(* IEC 61131-3 sources: daoli-st-library/DL_Process (part 35) *)

(* ---- FB_DL_FormationWeekPlan.st ---- *)
(*
  ==================================================================
  组件名 Component  : FB_DL_FormationWeekPlan
  分类   Category   : DL_Process
  版本   Version    : 1.0.0
  功能   Purpose    : 周计划窗（周序号闸 + 月窗闸双闸）。把日历日换算成「月内周
                      序号（1..5）」与「周内日序号（1..7）」，两个闸同时成立才算
                      计划窗开启：一 月窗闸 = 当日落在组态的月内生产窗区间；
                      二 周序号闸 = 当日所在周序号落在允许的周区间。
                      同时给出周内与月内剩余天数，供上层排产节拍使用。
  溯源   Origin     : 周序号 / 月窗双闸为通用排产窗语义；本件为 clean-room 实现，
                      仅借鉴来源分类与参数域组织（来源标签 roadmap-p2-weekplan），
                      道莅原创设计，未复制任何闭源代码行。
  平台   Platform   : 纯 IEC 61131-3（INT 整除与 MOD，除子为常量，无私有库）
  作者   Author     : 道莅代码库 · PLC 编程专家（R55）
  ------------------------------------------------------------------
  边界 Boundary     :
                      一 本件只判双闸与剩余天数，不生成工单、不判产量；
                      二 周序号按「月内第几周」口径（1 日为第 1 周第 1 日），非 ISO 周；
                      三 整除与取模的除子均为常量 7，且除前已把日序回钳到 1..31；
                      四 双闸任一不成立即关窗，关窗原因由两个独立布尔出口区分（R190）；
                      五 无全局变量、无外部变量声明、无物理地址寻址。
  输出契约 Output contract:
                      bMonthGateOk / bWeekGateOk 为两条独立闸的实时值，
                      bWindowOpen 仅在两条闸同时成立时为真（挂状态量）；
                      nWeekIdx 域 1..5，nDayInWeek 域 1..7，两者恒由回钳后的日序派生；
                      eCause 故障级成因与 bError 配对（R45），信息级永不置 bError。
  修订记录 Revision  :
    2026-11-20  v1.0.0  R55 首版（批 2 · 序号 9）
  ==================================================================
*)

TYPE E_DL_FwpCause :
(
    eNone       := 0,   // 无成因 / no cause
    eCfgIllegal := 1,   // 组态非法：年月日、窗界或周区间越域（故障级，与 bError 配对）/ illegal config, calendar, window bounds or week band out of domain
    eMonthGate  := 2,   // 月窗闸不成立（信息级）/ the monthly window gate does not hold, informational
    eWeekGate   := 3    // 周序号闸不成立（信息级）/ the week index gate does not hold, informational
);
END_TYPE

FUNCTION_BLOCK FB_DL_FormationWeekPlan
VAR_INPUT
    bEnable      : BOOL := TRUE;             // 使能，失能时关窗 [-] / enable, the window closes when disabled
    bReset       : BOOL := FALSE;           // 复位上升沿清故障锁存 [-] / reset rising edge clears the fault latch
    nYear        : INT := 2026;              // 当前年份 [年]，域 2000..2100 / current year [year], domain 2000 to 2100
    nMonth       : INT := 1;                 // 当前月份 [月]，域 1..12 / current month [month], domain 1 to 12
    nDayOfMonth  : INT := 1;                 // 当月第几日 [日]，域 1..31 / day of month [day], domain 1 to 31
    nWinStartDay : INT := 1;                 // 月生产窗起始日 [日] / monthly production window start day [day]
    nWinEndDay   : INT := 28;                // 月生产窗结束日 [日]，须不早于起始日 / monthly window end day, not earlier than the start
    nWeekFrom    : INT := 1;                 // 允许的周序号下限（月内第几周）[周]，域 1..5 / allowed week index floor, domain 1 to 5
    nWeekTo      : INT := 5;                 // 允许的周序号上限（月内第几周）[周]，域 1..5 / allowed week index ceiling, domain 1 to 5
END_VAR
VAR_OUTPUT
    bWindowOpen  : BOOL := FALSE;            // 双闸同时成立（计划窗开启）[-] / both gates hold, the planning window is open
    bMonthGateOk : BOOL := FALSE;            // 月窗闸实时值 [-] / monthly window gate live value
    bWeekGateOk  : BOOL := FALSE;            // 周序号闸实时值 [-] / week index gate live value
    nWeekIdx     : INT := 1;                 // 月内周序号 [周]，域 1..5 / week index within the month, domain 1 to 5
    nDayInWeek   : INT := 1;                 // 周内日序号 [日]，域 1..7 / day index within the week, domain 1 to 7
    nRemainInWeek: INT := 0;                 // 本周剩余天数（不跨月）[日] / remaining days this week, not crossing the month
    nRemainInMonth : INT := 0;               // 本月剩余天数 [日] / remaining days this month
    nPlanDays    : INT := 0;                 // 本窗剩余可排产天数（双闸内计数）[日] / remaining plannable days inside the window
    eCause       : E_DL_FwpCause := E_DL_FwpCause.eNone; // 成因出口 [枚举] / cause outlet [enum]
    bError       : BOOL := FALSE;            // 故障锁存标志 [-] / fault latch flag
END_VAR
VAR
    rtReset      : R_TRIG;                   // 复位沿检测，段 0 无条件刷新 / reset edge detector, refreshed unconditionally in segment zero
    _eFaultCause : E_DL_FwpCause := E_DL_FwpCause.eNone;  // 故障级成因，锁存至复位沿 / fault cause, latched until the reset edge
    _bFault      : BOOL := FALSE;            // 故障锁存位 [-] / fault latch bit
    _bInit       : BOOL := FALSE;            // 首扫初始化完成标志（R310）/ first scan initialisation flag
    _bCfgBad     : BOOL := FALSE;            // 组态非法判定 [-] / illegal configuration verdict
    _bMonthGate  : BOOL := FALSE;            // 月窗闸工作值 [-] / monthly window gate working value
    _bWeekGate   : BOOL := FALSE;            // 周序号闸工作值 [-] / week index gate working value
    _nDaysInMonth: INT := 30;                // 当月日历天数 [日] / calendar days of the current month [day]
    _nDay        : INT := 1;                 // 回钳后的当日序号 [日] / clamped day index [day]
    _nStart      : INT := 1;                 // 回钳后的窗起始日 [日] / clamped window start day [day]
    _nEnd        : INT := 1;                 // 回钳后的窗结束日 [日] / clamped window end day [day]
    _nWeekFrom   : INT := 1;                 // 回钳后的周序号下限 [周] / clamped week index floor [week]
    _nWeekTo     : INT := 5;                 // 回钳后的周序号上限 [周] / clamped week index ceiling [week]
    _nWeekIdx    : INT := 1;                 // 周序号工作值 [周] / week index working value [week]
    _nDayInWeek  : INT := 1;                 // 周内日序号工作值 [日] / day in week working value [day]
    _nRemainWeek : INT := 0;                 // 本周剩余天数工作值 [日] / remaining week days working value [day]
    _nRemainMonth: INT := 0;                 // 本月剩余天数工作值 [日] / remaining month days working value [day]
    _nPlanDays   : INT := 0;                 // 窗内剩余可排产天数工作值 [日] / remaining plannable days working value [day]
    _nScanDay    : INT := 1;                 // 窗内扫描用日序（自当日到窗末）[日] / scanning day index from today to the window end [day]
END_VAR
VAR CONSTANT
    DL_FWP_DAY_MAX   : INT := 31;            // 月内最大天数 [日] / maximum days within a month [day]
    DL_FWP_WEEK_N    : INT := 7;             // 一周日数，整除去子（常量非零）[日] / days per week, the division divisor as a non-zero constant [day]
    DL_FWP_WEEK_MAX  : INT := 5;             // 月内最大周序号 [周] / maximum week index within a month [week]
    DL_FWP_YEAR_MIN  : INT := 2000;          // 年份下限 [年] / year floor [year]
    DL_FWP_YEAR_MAX  : INT := 2100;          // 年份上限 [年] / year ceiling [year]
END_VAR

// 段 0｜复位沿无条件周期刷新（禁入分支）/ segment 0, unconditional refresh of the reset edge, never inside a branch
rtReset(CLK := bReset); // 复位沿无条件刷新 / unconditional refresh of the reset edge

// 段 1｜首扫初始化（R310）/ segment 1, first scan initialisation
IF NOT _bInit THEN // 首扫一拍 / the very first scan
    _bInit := TRUE; // 置首扫完成标志 / raise the first scan flag
    _bFault := FALSE; // 故障锁存清零 / clear the fault latch
    _eFaultCause := E_DL_FwpCause.eNone; // 故障级成因清零 / clear the fault cause
    _nWeekIdx := 1; // 周序号从第一周起 / the week index starts at one
    _nDayInWeek := 1; // 周内日序号从第一日起 / the day in week starts at one
END_IF

// 段 2｜复位沿作用域：清故障锁存与故障级成因（不动日历派生量）/ segment 2, reset edge scope
IF rtReset.Q THEN // 复位沿 / reset edge
    _bFault := FALSE; // 作用域一：清故障锁存 / scope one, clear the fault latch
    _eFaultCause := E_DL_FwpCause.eNone; // 作用域一：清故障级成因 / scope one, clear the fault cause
END_IF

// 段 3｜日历天数：闰年二月二十九日 / segment 3, calendar days with a leap February
_nDaysInMonth := 31; // 默认三十一日 / default thirty one days
CASE nMonth OF
1, 3, 5, 7, 8, 10, 12: // 大月 / long months
    _nDaysInMonth := 31; // 三十一日 / thirty one days
2: // 二月 / february
    IF ((nYear MOD 4) = 0) AND (((nYear MOD 100) <> 0) OR ((nYear MOD 400) = 0)) THEN // 闰年判据 / leap year criterion
        _nDaysInMonth := 29; // 闰年二十九日 / twenty nine days in a leap year
    ELSE
        _nDaysInMonth := 28; // 平年二十八日 / twenty eight days in a common year
    END_IF
4, 6, 9, 11: // 小月 / short months
    _nDaysInMonth := 30; // 三十日 / thirty days
ELSE // 非法月份兜底（R128）/ illegal month fallback
    _nDaysInMonth := 30; // 兜底三十日，故障另由域闸锁存 / fall back to thirty days, the fault is latched by the domain gate
END_CASE

// 段 4｜组态域闸（R151 全覆盖）/ segment 4, configuration domain gate over every pin
_bCfgBad := FALSE; // 组态非法预置假 / preset the illegal configuration verdict to false
IF (nYear < DL_FWP_YEAR_MIN) OR (nYear > DL_FWP_YEAR_MAX) THEN // 年份越域 / year out of domain
    _bCfgBad := TRUE; // 判非法 / mark illegal
END_IF
IF (nMonth < 1) OR (nMonth > 12) THEN // 月份越域 / month out of domain
    _bCfgBad := TRUE; // 判非法 / mark illegal
END_IF
IF (nDayOfMonth < 1) OR (nDayOfMonth > DL_FWP_DAY_MAX) THEN // 当日序号越域 / day index out of domain
    _bCfgBad := TRUE; // 判非法 / mark illegal
END_IF
IF (nWinStartDay < 1) OR (nWinStartDay > DL_FWP_DAY_MAX) OR (nWinEndDay < nWinStartDay) OR (nWinEndDay > DL_FWP_DAY_MAX) THEN // 窗界越域或自相矛盾 / window bounds out of domain or contradicting
    _bCfgBad := TRUE; // 判非法 / mark illegal
END_IF
IF (nWeekFrom < 1) OR (nWeekFrom > DL_FWP_WEEK_MAX) OR (nWeekTo < nWeekFrom) OR (nWeekTo > DL_FWP_WEEK_MAX) THEN // 周区间越域或自相矛盾 / week band out of domain or contradicting
    _bCfgBad := TRUE; // 判非法 / mark illegal
END_IF
IF _bCfgBad AND (NOT _bFault) THEN // 组态非法且未锁存 / illegal configuration and not yet latched
    _bFault := TRUE; // 置故障锁存 / raise the fault latch
    _eFaultCause := E_DL_FwpCause.eCfgIllegal; // 故障级成因 (R45 配对 bError) / fault grade cause paired with bError
END_IF

// 段 5｜回钳：日序、窗界、周区间一律回钳到可比较域 / segment 5, clamping the day, the window bounds and the week band
_nDay := nDayOfMonth; // 日序直通 / day index passes through
IF _nDay < 1 THEN // 下越界 / below the lower bound
    _nDay := 1; // 回钳到一日 / clamp to day one
ELSIF _nDay > _nDaysInMonth THEN // 上越界 / above the upper bound
    _nDay := _nDaysInMonth; // 回钳到月末 / clamp to the last day
END_IF
_nStart := nWinStartDay; // 窗起始日直通 / window start passes through
IF _nStart < 1 THEN // 下越界 / below the lower bound
    _nStart := 1; // 回钳到一日 / clamp to day one
ELSIF _nStart > _nDaysInMonth THEN // 上越界 / above the upper bound
    _nStart := _nDaysInMonth; // 回钳到月末 / clamp to the last day
END_IF
_nEnd := nWinEndDay; // 窗结束日直通 / window end passes through
IF _nEnd < _nStart THEN // 结束早于起始 / end earlier than start
    _nEnd := _nStart; // 回钳到起始日 / clamp to the start day
ELSIF _nEnd > _nDaysInMonth THEN // 上越界 / above the upper bound
    _nEnd := _nDaysInMonth; // 回钳到月末 / clamp to the last day
END_IF
_nWeekFrom := nWeekFrom; // 周下限直通 / the week floor passes through
IF _nWeekFrom < 1 THEN // 下越界 / below the lower bound
    _nWeekFrom := 1; // 回钳到第一周 / clamp to the first week
ELSIF _nWeekFrom > DL_FWP_WEEK_MAX THEN // 上越界 / above the upper bound
    _nWeekFrom := DL_FWP_WEEK_MAX; // 回钳到第五周 / clamp to the fifth week
END_IF
_nWeekTo := nWeekTo; // 周上限直通 / the week ceiling passes through
IF _nWeekTo < _nWeekFrom THEN // 上限早于下限 / ceiling earlier than the floor
    _nWeekTo := _nWeekFrom; // 回钳到下限 / clamp to the floor
ELSIF _nWeekTo > DL_FWP_WEEK_MAX THEN // 上越界 / above the upper bound
    _nWeekTo := DL_FWP_WEEK_MAX; // 回钳到第五周 / clamp to the fifth week
END_IF

// 段 6｜周序号与周内日序号派生：除子为常量 7，日序已回钳 1..31 / segment 6, week index and day in week derived with the constant divisor seven
_nWeekIdx := ((_nDay - 1) / DL_FWP_WEEK_N) + 1; // 月内周序号，整除除子为常量七 / week index within the month with the constant divisor seven
IF _nWeekIdx < 1 THEN // 下越界（防御）/ below the lower bound as a defence
    _nWeekIdx := 1; // 回钳到第一周 / clamp to the first week
ELSIF _nWeekIdx > DL_FWP_WEEK_MAX THEN // 上越界 / above the upper bound
    _nWeekIdx := DL_FWP_WEEK_MAX; // 回钳到第五周 / clamp to the fifth week
END_IF
_nDayInWeek := ((_nDay - 1) MOD DL_FWP_WEEK_N) + 1; // 周内日序，取模除子为常量七 / day in week with the constant divisor seven
IF _nDayInWeek < 1 THEN // 下越界（防御）/ below the lower bound as a defence
    _nDayInWeek := 1; // 回钳到第一日 / clamp to the first day
ELSIF _nDayInWeek > DL_FWP_WEEK_N THEN // 上越界 / above the upper bound
    _nDayInWeek := DL_FWP_WEEK_N; // 回钳到第七日 / clamp to the seventh day
END_IF

// 段 7｜双闸判定：月窗闸与周序号闸各自独立（R190 归因唯一）/ segment 7, the two gates evaluated independently
_bMonthGate := (_nDay >= _nStart) AND (_nDay <= _nEnd); // 月窗闸：当日落在月生产窗内 / monthly window gate
_bWeekGate := (_nWeekIdx >= _nWeekFrom) AND (_nWeekIdx <= _nWeekTo); // 周序号闸：周序号落在允许区间 / week index gate
IF NOT bEnable THEN // 失能：关窗（R191 显式声明）/ disabled, the window closes
    _bMonthGate := FALSE; // 月窗闸撤除 / the monthly gate is withdrawn
    _bWeekGate := FALSE; // 周序号闸撤除 / the week gate is withdrawn
END_IF

// 段 8｜剩余天数：周内剩余不跨月，窗内剩余按双闸逐日推演 / segment 8, remaining days within the week and inside the window
_nRemainWeek := DL_FWP_WEEK_N - _nDayInWeek; // 本周剩余天数（跨月部分由下一行截断）/ remaining days this week, truncated by the next line
IF (_nDay + _nRemainWeek) > _nDaysInMonth THEN // 周尾越过月末 / the week tail crosses the month end
    _nRemainWeek := _nDaysInMonth - _nDay; // 截断到月末 / truncated at the month end
END_IF
IF _nRemainWeek < 0 THEN // 防御：负值不可能 / defence, a negative value is impossible
    _nRemainWeek := 0; // 钳零 / clamped to zero
END_IF
_nRemainMonth := _nDaysInMonth - _nDay; // 本月剩余天数 / remaining days this month
IF _nRemainMonth < 0 THEN // 防御：负值不可能 / defence, a negative value is impossible
    _nRemainMonth := 0; // 钳零 / clamped to zero
END_IF
_nPlanDays := 0; // 窗内剩余可排产天数清零 / clear the remaining plannable days
IF _bMonthGate AND _bWeekGate THEN // 双闸内才逐日推演 / the day sweep only runs inside both gates
    _nScanDay := _nDay; // 自当日起扫 / sweep from today
    WHILE _nScanDay <= _nEnd DO // 扫到窗末为止，上界为回钳后的窗末日 / sweep up to the window end
        IF ((((_nScanDay - 1) / DL_FWP_WEEK_N) + 1) >= _nWeekFrom) AND ((((_nScanDay - 1) / DL_FWP_WEEK_N) + 1) <= _nWeekTo) THEN // 该日的周序号落在允许区间 / the week index of that day is inside the band
            _nPlanDays := _nPlanDays + 1; // 计入可排产天数 / count as a plannable day
        END_IF
        _nScanDay := _nScanDay + 1; // 日序递增 / increment the day index
    END_WHILE
END_IF

// 段 9｜成因分派（固定优先级：故障 > 月窗闸 > 周序号闸 > 无成因）/ segment 9, cause dispatch with a fixed priority
IF _bFault THEN // 故障锁存优先 / the fault latch takes priority
    eCause := _eFaultCause; // 故障级成因锁存回放 / the fault cause is replayed from the latch
ELSIF (NOT _bMonthGate) AND _bWeekGate THEN // 仅月窗闸不成立 / only the monthly gate fails
    eCause := E_DL_FwpCause.eMonthGate; // 信息级成因 / informational cause
ELSIF _bMonthGate AND (NOT _bWeekGate) THEN // 仅周序号闸不成立 / only the week gate fails
    eCause := E_DL_FwpCause.eWeekGate; // 信息级成因 / informational cause
ELSIF (NOT _bMonthGate) AND (NOT _bWeekGate) THEN // 两闸均不成立 / both gates fail
    eCause := E_DL_FwpCause.eMonthGate; // 按月窗闸优先报告（上游先解除大闸）/ report the monthly gate first because the upstream gate must clear first
ELSE
    eCause := E_DL_FwpCause.eNone; // 双闸内无成因 / no cause inside both gates
END_IF

// 段 10｜统一出口 / segment 10, unified outlet
bMonthGateOk := _bMonthGate; // 月窗闸出口 / monthly gate outlet
bWeekGateOk := _bWeekGate; // 周序号闸出口 / week gate outlet
bWindowOpen := _bMonthGate AND _bWeekGate; // 双闸合成（挂状态量，非单拍标志）/ the composite gate as a state quantity
nWeekIdx := _nWeekIdx; // 周序号出口 / week index outlet
nDayInWeek := _nDayInWeek; // 周内日序号出口 / day in week outlet
nRemainInWeek := _nRemainWeek; // 本周剩余天数出口 / remaining week days outlet
nRemainInMonth := _nRemainMonth; // 本月剩余天数出口 / remaining month days outlet
nPlanDays := _nPlanDays; // 窗内可排产天数出口 / remaining plannable days outlet
bError := _bFault; // 故障标志与锁存位同源 / the fault flag shares the latch source
END_FUNCTION_BLOCK

(* ---- FB_DL_FormatMonthAudit.st ---- *)
(*
  ==================================================================
  组件名 Component  : FB_DL_FormatMonthAudit
  分类   Category   : DL_Process
  版本   Version    : 1.0.0
  功能   Purpose    : 化成 / 分容月度窗排产审计。按日历日判月度生产窗是否开启，
                      窗内以「已完数量 / 月计划数量」与「窗内已过比例」两条进度
                      比对，给出准时 / 落后 / 超前三种审计结论，并在窗关闭那一拍
                      输出审计收口脉冲与收口结论（结论锁存至下月开窗）。
  溯源   Origin     : 月度窗进度审计为通用排产审计语义；本件为 clean-room 实现，
                      仅借鉴来源分类与参数域组织（来源标签 roadmap-p2-formation），
                      道莅原创设计，未复制任何闭源代码行。
  平台   Platform   : 纯 IEC 61131-3（R_TRIG / REAL / UDINT 运算，无私有库）
  作者   Author     : 道莅代码库 · PLC 编程专家（R55）
  ------------------------------------------------------------------
  边界 Boundary     :
                      一 本件只做审计判级与收口脉冲，不派工单、不改计划量（属主边界）；
                      二 窗内已过比例按「窗首日至当日」计，窗关闭后比例钳到 100%；
                      三 计划量为零判组态故障并锁存至复位沿，不做除法；
                      四 数量类走 UDINT 直比（禁 ABS 单侧判越界，R55 口径）；
                      五 无全局变量、无外部变量声明、无物理地址寻址。
  输出契约 Output contract:
                      eAudit 四态互斥（eNone 仅在窗关闭或未参与时出现）；
                      bAuditClose 为单拍脉冲（内部位置位、统一出口映射后撤销）；
                      fCompletePct / fReqDailyRate 在除子不可用时保持上拍值；
                      eCause 故障级成因与 bError 配对（R45），信息级永不置 bError。
  修订记录 Revision  :
    2026-11-20  v1.0.0  R55 首版（批 2 · 序号 6）
  ==================================================================
*)

TYPE E_DL_FmaAudit :
(
    eNone    := 0,      // 无结论：窗未开或已收口 / no verdict, the window is closed or not yet opened
    eOnPlan  := 10,     // 准时：实际进度落在期望带内 / on plan, the actual progress sits inside the expected band
    eBehind  := 20,     // 落后：实际进度低于期望带下沿 / behind, the actual progress is below the band
    eAhead   := 30      // 超前：实际进度高于期望带上沿 / ahead, the actual progress is above the band
);
END_TYPE

TYPE E_DL_FmaCause :
(
    eNone       := 0,   // 无成因 / no cause
    eCfgIllegal := 1,   // 组态非法：年月日或窗界越域（故障级，与 bError 配对）/ illegal config, calendar or window bounds out of domain
    ePlanZero   := 2,   // 月计划量为零，进度不可算（故障级，与 bError 配对）/ monthly plan is zero, progress not computable
    eWinClosed  := 3    // 当前不在生产窗内（信息级）/ the current day is outside the production window, informational
);
END_TYPE

FUNCTION_BLOCK FB_DL_FormatMonthAudit
VAR_INPUT
    bEnable      : BOOL := TRUE;             // 使能，失能时结论冻结保持 [-] / enable, the verdict freezes and holds when disabled
    bReset       : BOOL := FALSE;           // 复位上升沿清故障锁存与收口结论 [-] / reset rising edge clears the fault latch and the closing verdict
    nYear        : INT := 2026;              // 当前年份 [年]，域 2000..2100 / current year [year], domain 2000 to 2100
    nMonth       : INT := 1;                 // 当前月份 [月]，域 1..12 / current month [month], domain 1 to 12
    nDayOfMonth  : INT := 1;                 // 当月第几日 [日]，域 1..31 / day of month [day], domain 1 to 31
    nWinStartDay : INT := 1;                 // 生产窗起始日 [日] / production window start day [day]
    nWinEndDay   : INT := 25;                // 生产窗结束日 [日]，须不早于起始日 / production window end day, not earlier than the start
    uPlanCells   : UDINT := 1000;            // 月度计划数量 [只]，域 大于零 / monthly planned quantity [pieces], domain above zero
    uDoneCells   : UDINT := 0;               // 已完数量 [只] / completed quantity [pieces]
    fBehindPct   : REAL := 5.0;              // 落后判定带宽度 [百分比]，域 大于零 / behind band width [percent], domain above zero
    fAheadPct    : REAL := 10.0;             // 超前判定带宽度 [百分比]，域 大于零 / ahead band width [percent], domain above zero
END_VAR
VAR_OUTPUT
    bWindowOpen  : BOOL := FALSE;            // 生产窗是否开启 [-] / production window open flag
    nRemainDays  : INT := 0;                 // 窗内剩余天数（窗关闭为 0）[日] / remaining window days, zero when closed
    nElapsedDays : INT := 0;                 // 窗内已过天数（含当日）[日] / elapsed window days including today
    fCompletePct : REAL := 0.0;              // 实际完成比例 [百分比] / actual completion ratio [percent]
    fExpectPct   : REAL := 0.0;              // 按时进度期望比例 [百分比] / expected on-time progress ratio [percent]
    fReqDailyRate: REAL := 0.0;              // 达产所需日均量 [只每日] / required daily rate to hit the plan [pieces per day]
    eAudit       : E_DL_FmaAudit := E_DL_FmaAudit.eNone; // 审计结论出口 [枚举] / audit verdict outlet [enum]
    eAuditClose  : E_DL_FmaAudit := E_DL_FmaAudit.eNone; // 窗关闭拍锁存的收口结论 [枚举] / verdict latched at window closing [enum]
    bAuditClose  : BOOL := FALSE;            // 审计收口单拍脉冲 [-] / audit closing single-shot pulse
    eCause       : E_DL_FmaCause := E_DL_FmaCause.eNone; // 成因出口 [枚举] / cause outlet [enum]
    bError       : BOOL := FALSE;            // 故障锁存标志 [-] / fault latch flag
END_VAR
VAR
    rtReset      : R_TRIG;                   // 复位沿检测，段 0 无条件刷新 / reset edge detector, refreshed unconditionally in segment zero
    _eCause      : E_DL_FmaCause := E_DL_FmaCause.eNone;   // 信息级成因，每拍重算 / informational cause, recomputed every scan
    _eFaultCause : E_DL_FmaCause := E_DL_FmaCause.eNone;   // 故障级成因，锁存至复位沿 / fault cause, latched until the reset edge
    _eAudit      : E_DL_FmaAudit := E_DL_FmaAudit.eNone;   // 内部结论 / internal verdict
    _eAuditClose : E_DL_FmaAudit := E_DL_FmaAudit.eNone;   // 收口结论锁存 / latched closing verdict
    _bFault      : BOOL := FALSE;            // 故障锁存位 [-] / fault latch bit
    _bInit       : BOOL := FALSE;            // 首扫初始化完成标志（R310）/ first scan initialisation flag
    _bWinOpenPrev: BOOL := FALSE;            // 上一拍窗开启快照，收口沿判据用 [-] / previous scan window flag for the closing edge
    _bCloseInt   : BOOL := FALSE;            // 收口脉冲内部位，统一出口映射 / internal closing pulse bit, mapped at the unified outlet
    _bWinOpen    : BOOL := FALSE;            // 本拍窗开启判定 [-] / this scan window open verdict
    _bCfgBad     : BOOL := FALSE;            // 组态非法判定 [-] / illegal configuration verdict
    _bDivOk      : BOOL := FALSE;            // 除子可用判定（计划量非零）[-] / divisor usable verdict
    _nDaysInMonth: INT := 30;                // 当月日历天数 [日] / calendar days of the current month [day]
    _nStart      : INT := 1;                 // 钳定后的窗起始日 [日] / clamped window start day [day]
    _nEnd        : INT := 1;                 // 钳定后的窗结束日 [日] / clamped window end day [day]
    _nDay        : INT := 1;                 // 钳定后的当日序号 [日] / clamped day index [day]
    _nElapsed    : INT := 0;                 // 窗内已过天数工作值 [日] / elapsed window days working value [day]
    _nRemain     : INT := 0;                 // 窗内剩余天数工作值 [日] / remaining window days working value [day]
    _nWinLen     : INT := 1;                 // 窗长（天数）[日] / window length in days [day]
    _fPlan       : REAL := 0.0;              // 计划量实数化暂存 [只] / planned quantity as a real [pieces]
    _fDone       : REAL := 0.0;              // 已完量实数化暂存 [只] / completed quantity as a real [pieces]
    _fComplete   : REAL := 0.0;              // 完成比例工作值 [百分比] / completion ratio working value [percent]
    _fExpect     : REAL := 0.0;              // 期望比例工作值 [百分比] / expected ratio working value [percent]
    _fReqRate    : REAL := 0.0;              // 所需日均量工作值 [只每日] / required daily rate working value [pieces per day]
    _fGap        : REAL := 0.0;              // 计划缺口 [只] / remaining plan gap [pieces]
    _fDivWin     : REAL := 1.0;              // 窗长除子 [日]，已证不小于 1 / window length divisor proven not below one
    _fDivDay     : REAL := 1.0;              // 剩余天数除子 [日]，已证不小于 1 / remaining day divisor proven not below one
END_VAR
VAR CONSTANT
    DL_FMA_DAY_MAX   : INT := 31;            // 月内最大天数 [日] / maximum days within a month [day]
    DL_FMA_YEAR_MIN  : INT := 2000;          // 年份下限 [年] / year floor [year]
    DL_FMA_YEAR_MAX  : INT := 2100;          // 年份上限 [年] / year ceiling [year]
    DL_FMA_BAND_MAX  : REAL := 100.0;        // 判定带宽度上限 [百分比] / band width ceiling [percent]
    DL_FMA_PCT_MAX   : REAL := 1000.0;       // 完成比例上限，防计划量过小放大 [百分比] / completion ratio ceiling against a tiny plan
    DL_FMA_RATE_MAX  : REAL := 1.0E7;        // 日均量上限，防除子过小放大 [只每日] / daily rate ceiling against a tiny divisor
END_VAR

// 段 0｜复位沿无条件周期刷新（禁入分支）/ segment 0, unconditional refresh of the reset edge, never inside a branch
rtReset(CLK := bReset); // 复位沿无条件刷新 / unconditional refresh of the reset edge

// 段 1｜首扫初始化（R310）/ segment 1, first scan initialisation
IF NOT _bInit THEN // 首扫一拍 / the very first scan
    _bInit := TRUE; // 置首扫完成标志 / raise the first scan flag
    _bFault := FALSE; // 故障锁存清零 / clear the fault latch
    _eCause := E_DL_FmaCause.eNone; // 信息级成因清零 / clear the informational cause
    _eFaultCause := E_DL_FmaCause.eNone; // 故障级成因清零 / clear the fault cause
    _eAudit := E_DL_FmaAudit.eNone; // 结论清零 / clear the verdict
    _eAuditClose := E_DL_FmaAudit.eNone; // 收口结论清零 / clear the closing verdict
    _bWinOpenPrev := FALSE; // 窗开启快照清零 / clear the window snapshot
END_IF

// 段 2｜复位沿作用域：清故障锁存 / 清收口结论 / 清窗快照（结论不改，避免审计断档）/ segment 2, reset edge scope
IF rtReset.Q THEN // 复位沿 / reset edge
    _bFault := FALSE; // 作用域一：清故障锁存 / scope one, clear the fault latch
    _eFaultCause := E_DL_FmaCause.eNone; // 作用域一：清故障级成因 / scope one, clear the fault cause
    _eAuditClose := E_DL_FmaAudit.eNone; // 作用域二：清收口结论 / scope two, clear the closing verdict
    _bCloseInt := FALSE; // 作用域二：清收口脉冲内部位 / scope two, clear the internal closing bit
    _bWinOpenPrev := FALSE; // 作用域三：清窗开启快照 / scope three, clear the window snapshot
END_IF

// 段 3｜日历天数：闰年二月二十九日，其余按大小月 / segment 3, calendar days with a leap February
_nDaysInMonth := 31; // 默认三十一日 / default thirty one days
CASE nMonth OF
1, 3, 5, 7, 8, 10, 12: // 大月 / long months
    _nDaysInMonth := 31; // 三十一日 / thirty one days
2: // 二月 / february
    IF ((nYear MOD 4) = 0) AND (((nYear MOD 100) <> 0) OR ((nYear MOD 400) = 0)) THEN // 闰年判据 / leap year criterion
        _nDaysInMonth := 29; // 闰年二十九日 / twenty nine days in a leap year
    ELSE
        _nDaysInMonth := 28; // 平年二十八日 / twenty eight days in a common year
    END_IF
4, 6, 9, 11: // 小月 / short months
    _nDaysInMonth := 30; // 三十日 / thirty days
ELSE // 非法月份兜底（R128）/ illegal month fallback
    _nDaysInMonth := 30; // 兜底三十日，故障另由域闸锁存 / fall back to thirty days, the fault is latched by the domain gate
END_CASE

// 段 4｜组态域闸（R151 全覆盖）：年月日、窗界、计划量、判定带 / segment 4, configuration domain gate over every pin
_bCfgBad := FALSE; // 组态非法预置假 / preset the illegal configuration verdict to false
IF (nYear < DL_FMA_YEAR_MIN) OR (nYear > DL_FMA_YEAR_MAX) THEN // 年份越域 / year out of domain
    _bCfgBad := TRUE; // 判非法 / mark illegal
END_IF
IF (nMonth < 1) OR (nMonth > 12) THEN // 月份越域 / month out of domain
    _bCfgBad := TRUE; // 判非法 / mark illegal
END_IF
IF (nDayOfMonth < 1) OR (nDayOfMonth > DL_FMA_DAY_MAX) THEN // 当日序号越域 / day index out of domain
    _bCfgBad := TRUE; // 判非法 / mark illegal
END_IF
IF (nWinStartDay < 1) OR (nWinStartDay > DL_FMA_DAY_MAX) OR (nWinEndDay < nWinStartDay) OR (nWinEndDay > DL_FMA_DAY_MAX) THEN // 窗界越域或自相矛盾 / window bounds out of domain or contradicting
    _bCfgBad := TRUE; // 判非法 / mark illegal
END_IF
IF (fBehindPct <= 0.0) OR (fBehindPct > DL_FMA_BAND_MAX) OR (fBehindPct <> fBehindPct) THEN // 落后带宽越域 / behind band out of domain
    _bCfgBad := TRUE; // 判非法 / mark illegal
END_IF
IF (fAheadPct <= 0.0) OR (fAheadPct > DL_FMA_BAND_MAX) OR (fAheadPct <> fAheadPct) THEN // 超前带宽越域 / ahead band out of domain
    _bCfgBad := TRUE; // 判非法 / mark illegal
END_IF
IF _bCfgBad AND (NOT _bFault) THEN // 组态非法且未锁存 / illegal configuration and not yet latched
    _bFault := TRUE; // 置故障锁存 / raise the fault latch
    _eFaultCause := E_DL_FmaCause.eCfgIllegal; // 故障级成因 (R45 配对 bError) / fault grade cause paired with bError
END_IF

// 段 5｜钳定：窗界与当日一律回钳到当月日历范围内（回钳后可安全比较）/ segment 5, clamping the window bounds and the day into the calendar range
_nStart := nWinStartDay; // 窗起始日直通 / window start passes through
IF _nStart < 1 THEN // 下越界 / below the lower bound
    _nStart := 1; // 回钳到一日 / clamp to day one
ELSIF _nStart > _nDaysInMonth THEN // 上越界 / above the upper bound
    _nStart := _nDaysInMonth; // 回钳到月末 / clamp to the last day
END_IF
_nEnd := nWinEndDay; // 窗结束日直通 / window end passes through
IF _nEnd < _nStart THEN // 结束早于起始 / end earlier than start
    _nEnd := _nStart; // 回钳到起始日，窗长退化为一日 / clamp to the start so the window degenerates to a single day
ELSIF _nEnd > _nDaysInMonth THEN // 上越界 / above the upper bound
    _nEnd := _nDaysInMonth; // 回钳到月末 / clamp to the last day
END_IF
_nDay := nDayOfMonth; // 当日序号直通 / day index passes through
IF _nDay < 1 THEN // 下越界 / below the lower bound
    _nDay := 1; // 回钳到一日 / clamp to day one
ELSIF _nDay > _nDaysInMonth THEN // 上越界 / above the upper bound
    _nDay := _nDaysInMonth; // 回钳到月末 / clamp to the last day
END_IF

// 段 6｜窗开启与窗内已过 / 剩余天数 / segment 6, window open verdict with elapsed and remaining days
_nWinLen := _nEnd - _nStart + 1; // 窗长（闭区间）[日] / window length over a closed interval [day]
IF _nWinLen < 1 THEN // 窗长为零不可能（已回钳）/ a zero length is impossible after clamping
    _nWinLen := 1; // 兜底一日，防除零 / fall back to one against division by zero
END_IF
_bWinOpen := (_nDay >= _nStart) AND (_nDay <= _nEnd); // 窗开启判据 / window open criterion
IF _bWinOpen THEN // 窗内 / inside the window
    _nElapsed := _nDay - _nStart + 1; // 已过天数含当日 / elapsed days including today
    _nRemain := _nEnd - _nDay; // 剩余天数不含当日 / remaining days excluding today
ELSE // 窗外 / outside the window
    _nElapsed := 0; // 已过天数零 / elapsed days zero
    _nRemain := 0; // 剩余天数零 / remaining days zero
END_IF
IF NOT bEnable THEN // 失能：结论与比例冻结保持末值（R191 显式声明）/ disabled, ratios and verdict freeze and hold their last value
    _bWinOpen := FALSE; // 窗开启标志撤除 / the window flag is withdrawn
END_IF

// 段 7｜比例与日均：计划量为零不计算，除子先域闸 / segment 7, ratios and daily rate with both divisors gated first
_bDivOk := uPlanCells > 0; // 计划量非零才可算比例 / the plan must be non-zero for any ratio
_eCause := E_DL_FmaCause.eNone; // 信息级成因每拍重算（R190 归因唯一）/ the informational cause is recomputed every scan
IF NOT _bDivOk THEN // 计划量为零 / the plan is zero
    IF NOT _bFault THEN // 未锁存才记故障 / record the fault only when not yet latched
        _bFault := TRUE; // 置故障锁存 / raise the fault latch
        _eFaultCause := E_DL_FmaCause.ePlanZero; // 故障级成因 (R45 配对 bError) / fault grade cause paired with bError
    END_IF
END_IF
IF _bDivOk AND _bWinOpen THEN // 计划可用且在窗内 / the plan is usable and the window is open
    _fPlan := UDINT_TO_REAL(uPlanCells); // 计划量实数化 / planned quantity as a real
    _fDone := UDINT_TO_REAL(uDoneCells); // 已完量实数化 / completed quantity as a real
    _fComplete := _fDone / _fPlan * 100.0; // 完成比例，除子已证大于零 / completion ratio, divisor proven positive
    IF _fComplete > DL_FMA_PCT_MAX THEN // 比例越上限 / ratio above the ceiling
        _fComplete := DL_FMA_PCT_MAX; // 上钳，防计划量过小放大 / clamp upward against a tiny plan
    END_IF
    _fDivWin := INT_TO_REAL(_nWinLen); // 窗长除子，已证不小于 1 / window length divisor proven not below one
    _fExpect := INT_TO_REAL(_nElapsed) / _fDivWin * 100.0; // 期望比例 / expected ratio
    _fGap := _fPlan - _fDone; // 计划缺口 / plan gap
    IF _fGap < 0.0 THEN // 已完成超出计划 / the plan is already exceeded
        _fGap := 0.0; // 缺口归零 / gap zeroed
    END_IF
    IF _nRemain > 0 THEN // 有剩余天数 / remaining days exist
        _fDivDay := INT_TO_REAL(_nRemain); // 剩余天数除子，已证大于零 / remaining day divisor proven positive
        _fReqRate := _fGap / _fDivDay; // 所需日均量 / required daily rate
        IF _fReqRate > DL_FMA_RATE_MAX THEN // 日均量越上限 / daily rate above the ceiling
            _fReqRate := DL_FMA_RATE_MAX; // 上钳，防除子过小放大 / clamp upward against a tiny divisor
        END_IF
    ELSE // 无剩余天数（窗末日或窗关闭）/ no remaining days
        _fReqRate := 0.0; // 日均需求归零 / the daily requirement is zeroed
    END_IF
    IF (_fComplete < (_fExpect - fBehindPct)) THEN // 实际低于期望带下沿 / actual below the band
        _eAudit := E_DL_FmaAudit.eBehind; // 判落后 / behind verdict
    ELSIF (_fComplete > (_fExpect + fAheadPct)) THEN // 实际高于期望带上沿 / actual above the band
        _eAudit := E_DL_FmaAudit.eAhead; // 判超前 / ahead verdict
    ELSE // 落在带内 / inside the band
        _eAudit := E_DL_FmaAudit.eOnPlan; // 判准时 / on plan verdict
    END_IF
ELSIF _bDivOk THEN // 计划可用但窗外 / the plan is usable yet outside the window
    _eAudit := E_DL_FmaAudit.eNone; // 窗外无结论 / no verdict outside the window
    _eCause := E_DL_FmaCause.eWinClosed; // 信息级成因：不在窗内 / informational cause, outside the window
END_IF

// 段 8｜收口沿：上一拍在窗内、本拍在窗外 → 锁存结论并出单拍脉冲 / segment 8, closing edge latches the verdict and raises a single-shot pulse
IF _bWinOpenPrev AND (NOT _bWinOpen) THEN // 窗关闭沿 / window closing edge
    _eAuditClose := _eAudit; // 结论锁存（窗内最后一拍的判级）/ latch the verdict from the last in-window scan
    IF _eAuditClose = E_DL_FmaAudit.eNone THEN // 收口拍无有效判级 / no valid verdict at closing
        _eAuditClose := E_DL_FmaAudit.eBehind; // 无结论按落后处理（保守侧，安全方向）/ no verdict is treated as behind on the conservative side
    END_IF
    _bCloseInt := TRUE; // 收口脉冲内部位置位（统一出口映射，R187）/ raise the internal pulse bit, mapped at the unified outlet
END_IF
_bWinOpenPrev := _bWinOpen; // 窗开启快照推进 / advance the window snapshot

// 段 9｜统一出口 / segment 9, unified outlet
bWindowOpen := _bWinOpen; // 窗开启出口 / window open outlet
nRemainDays := _nRemain; // 剩余天数出口 / remaining days outlet
nElapsedDays := _nElapsed; // 已过天数出口 / elapsed days outlet
fCompletePct := _fComplete; // 完成比例出口 / completion ratio outlet
fExpectPct := _fExpect; // 期望比例出口 / expected ratio outlet
fReqDailyRate := _fReqRate; // 所需日均量出口 / required daily rate outlet
eAudit := _eAudit; // 结论出口单点映射 / single-point verdict outlet mapping
eAuditClose := _eAuditClose; // 收口结论出口（锁存量）/ closing verdict outlet from the latch
bAuditClose := _bCloseInt; // 收口脉冲映射本拍值 / map the closing pulse for this scan
_bCloseInt := FALSE; // 映射后立即撤销，保证单拍宽度（R187 两段式）/ revoke right after mapping to keep a single-scan width
IF _bFault THEN // 故障锁存优先 / the fault latch takes priority
    eCause := _eFaultCause; // 故障级成因锁存回放 / the fault cause is replayed from the latch
ELSE
    eCause := _eCause; // 信息级成因直映 / the informational cause is mapped directly
END_IF
bError := _bFault; // 故障标志与锁存位同源 / the fault flag shares the latch source
END_FUNCTION_BLOCK

(* ---- FB_DL_FoupRfidCheck.st ---- *)
(*==============================================================================
 * 组件名称 (Component)  : FB_DL_FoupRfidCheck
 * 所属子库 (Sublibrary) : DL_Process
 * 当前版本 (Version)    : 1.0.0
 * 兼容性   (Platform)   : CODESYS 3.5+ / TwinCAT 3 / 汇川 InoProShop / 施耐德 Machine Expert
 *                         仅依赖 Standard.library（TON / R_TRIG / LEN），零厂商私有库
 * 功能描述 (Function)   : FOUP 身份校验与配方放行。
 *                         装载口读 FOUP 身份码后，按**固定顺序的四段校验链**裁决是否放行加工：
 *                           ① 身份码非空（空码 = 没读到，不放行）；
 *                           ② 身份码长度在 [uIdMinLen, uIdMaxLen] 内（格式闸，防半截码/粘码）；
 *                           ③ 在机配方非空（无配方不许放行）；
 *                           ④ 在机配方 = 期望配方（配方一致性，逐字符比对）。
 *                         四段任一失败即锁存失败原因，**且首因不覆盖**：第一个失败段决定 eCause，
 *                         后续段不再改写（R190 归因唯一）；放行在四段全过时才给单拍脉冲。
 *                         验收向量：
 *                           ① FOUP='F0012'，配方 'RCP-A' = 期望 'RCP-A' → bPass 单拍
 *                           ② FOUP=''                              → eIdEmpty 锁存
 *                           ③ FOUP='F01'（长度 < 4）                → eIdFormat 锁存
 *                           ④ 配方 'RCP-B' ≠ 期望 'RCP-A'          → eRecipeMismatch 锁存
 *                           ⑤ 启动后 tReadTo 内无读码完成             → eReadTimeout 锁存
 * 接口     (Interface)  : 入 bStartCheck 校验启动沿、bReadDone 读码完成沿、sFoupId FOUP 身份码、
 *                         sRecipeId 在机配方号、sExpectedRecipe 期望配方号、uIdMinLen / uIdMaxLen
 *                         身份码长度域、tReadTo 读码超时、bReset 复位沿；
 *                         出 bPass 放行脉冲（单拍）、bCheckFailed 校验失败锁存、bWaiting 等读码中、
 *                         eState 相、eCause 成因、bError 故障标志。
 * 边界     (Boundary)   : ① **属主边界（写死）：本件只做"身份 + 配方"校验链与放行脉冲，
 *                         不驱动装载口门/夹紧、不切配方、不写 MES 账**（分别属门件、配方件、通讯件）；
 *                         ② **长度域闸**：uIdMinLen ≥ 1 且 uIdMaxLen ≥ uIdMinLen 且 uIdMaxLen ≤ 15，
 *                         违反即锁存 eCfgIllegal（长度域非法会让格式闸静默失效，R179）；
 *                         ③ **超时 TON 冻结**：tonRead 的 IN 串 (NOT _bFault)，故障期不累计，
 *                         复位同拍不会立即重锁（R252）；TON 段 0 无条件调用；
 *                         ④ **锁存解除式**：bCheckFailed 与 eFault 仅由 bReset 上升沿解除
 *                         （R228B 唯一迁出）；bReset 为外部引脚、恒可达；
 *                         ⑤ **等待相退出条件 ≥2**：读码完成沿 ∨ 超时（R98/R129），
 *                         并补一条"启动命令已撤销 → 回待机"（进相前置消失出口）；
 *                         ⑥ 零全局耦合、零物理地址。
 * 分工声明 (Scope)      : 本件只管"FOUP 身份与配方放行校验"。不接管：载具路径路由
 *                         （属 FB_DL_RfidTrayRoute）、配方参数下发与切换（属配方件）、
 *                         FOUP 内部晶圆计数校验（属片盒件）。
 * 来源标签 (Source Tag) : ROADMAP 空勾真缺口 P1（FOUP 配方放行，自研 clean-room）
 * 码表     (Codes)      : 本件不占用任何全局数字码位（零码位范式 R297）；诊断由 BOOL + ENUM 出口承担。
 * 红线自检 (Redline)    : R1 ✓ 零 GVL/VAR_EXTERNAL ｜ R2 ✓ 零 %I/%Q/%M ｜ R3 ✓ 纯 IEC 61131-3
 *                         R4 ✓ 长度域闸 + 空串闸 + 超时 + 等待相双出口 ｜ R5 ✓ 声明逐行同行双语注释
 *                         R6 ✓ ENUM+CASE 含 ELSE 兜底 ｜ R7 ✓ TON/R_TRIG 段 0 无条件刷新
 * 修订历史 (Revision)   : 2026-11-19  v1.0.0  R47 首版（批次 3 · 序号 12）
 *==============================================================================*)

TYPE E_DL_FrcState :
(
    eIdle  := 0,    // 待机相（等校验启动） / Idle, awaiting a check request
    eWait  := 10,   // 等读码相（读码窗内） / Waiting for the tag read
    eFault := 90    // 故障相（等复位） / Fault, awaiting reset
);
END_TYPE

TYPE E_DL_FrcCause :
(
    eNone          := 0,   // 无异常 / No anomaly
    eIdEmpty       := 1,   // 身份码空（锁存） / Empty identity, latched
    eIdFormat      := 2,   // 身份码长度越域（锁存） / Identity length out of range, latched
    eRecipeEmpty   := 3,   // 在机配方空（锁存） / Empty on-machine recipe, latched
    eRecipeMismatch:= 4,   // 配方不一致（锁存） / Recipe mismatch, latched
    eReadTimeout   := 5,   // 读码超时（锁存） / Read timeout, latched
    eCfgIllegal    := 6,   // 组态非法（长度域/超时越域） / Illegal configuration
    ePhaseBad      := 7    // 非法相位兜底 / Illegal phase fallback
);
END_TYPE

FUNCTION_BLOCK FB_DL_FoupRfidCheck
VAR_INPUT
    bStartCheck    : BOOL := FALSE;      // 校验启动沿 [-] / Check-start edge
    bReadDone      : BOOL := FALSE;      // 读码完成沿 [-] / Tag-read edge
    sFoupId        : STRING[15] := '';   // FOUP 身份码（≤15 字符） [-] / FOUP identity, up to 15 chars
    sRecipeId      : STRING[15] := '';   // 在机配方号 [-] / On-machine recipe identifier
    sExpectedRecipe: STRING[15] := '';   // 期望配方号 [-] / Expected recipe identifier
    uIdMinLen      : UINT := 4;          // 身份码最小长度，域 1..15 [字符] / Minimum identity length
    uIdMaxLen      : UINT := 15;         // 身份码最大长度，域 ≥ 最小长度 [字符] / Maximum identity length
    tReadTo        : TIME := T#5S;       // 读码超时，域 > T#0S [ms] / Read timeout, > T#0S
    bReset         : BOOL := FALSE;      // 故障复位沿 [-] / Fault reset edge
END_VAR
VAR_OUTPUT
    bPass       : BOOL := FALSE;                         // 放行脉冲（单拍，四段全过） [-] / Pass pulse, single scan
    bCheckFailed: BOOL := FALSE;                         // 校验失败锁存（等复位） [-] / Check failure, latched
    bWaiting    : BOOL := FALSE;                         // 等读码中 [-] / Waiting for the tag read
    eState      : E_DL_FrcState := E_DL_FrcState.eIdle;  // 相出口 [-] / Phase outlet
    eCause      : E_DL_FrcCause := E_DL_FrcCause.eNone;  // 成因出口（R190 归因唯一） [-] / Cause outlet
    bError      : BOOL := FALSE;                         // 故障标志（仅故障级成因） [-] / Error flag, fault level only
END_VAR
VAR
    _eState   : E_DL_FrcState := E_DL_FrcState.eIdle;    // 内部相（CASE 唯一写入目标） / Internal phase
    _eCause   : E_DL_FrcCause := E_DL_FrcCause.eNone;    // 成因锁存量 / Latched cause
    _bFault   : BOOL := FALSE;                           // 故障锁存位 / Latched fault bit
    _bFail    : BOOL := FALSE;                           // 校验失败锁存位 / Latched check-failure bit
    _bPass    : BOOL := FALSE;                           // 放行脉冲内部位（单拍） / Internal pass pulse
    _bCfgBad  : BOOL := FALSE;                           // 组态非法当拍量 / Illegal configuration this scan
    _iLen     : INT := 0;                                // 身份码实际长度 [字符] / Actual identity length
    tonRead   : TON;                                     // 读码超时实例，段 0 无条件调用 / Read timeout instance
    rtStart   : R_TRIG;                                  // 启动沿实例，段 0 无条件调用 / Start edge instance
    rtRead    : R_TRIG;                                  // 读码沿实例，段 0 无条件调用 / Read edge instance
    rtReset   : R_TRIG;                                  // 复位沿实例，段 0 无条件调用 / Reset edge instance
END_VAR
VAR CONSTANT
    DL_FRC_LEN_MAX : UINT := 15;         // 身份码长度硬上限（与 STRING[15] 同源） [字符] / Hard length ceiling
END_VAR

(* —— 段 0：组态闸 + TON 与三沿无条件周期刷新（R228A；IN 串故障否决，R252） —— *)
_bCfgBad := (uIdMinLen < 1) OR (uIdMaxLen < uIdMinLen) OR (uIdMaxLen > DL_FRC_LEN_MAX)   // 长度域须满足 1 ≤ min ≤ max ≤ 15
         OR (tReadTo <= T#0S);                                                             // 超时须为正
rtStart(CLK := bStartCheck);                                                               // 启动沿 / Start edge
rtRead(CLK := bReadDone);                                                                  // 读码沿 / Read edge
rtReset(CLK := bReset);                                                                    // 复位沿 / Reset edge
tonRead(IN := (_eState = E_DL_FrcState.eWait) AND (NOT _bFault), PT := tReadTo);            // 读码超时（等读码相派生） / Read timeout

(* —— 段 1：单拍量预清零（锁存量 _eCause/_bFault/_bFail 不入清单，R107） —— *)
_bPass := FALSE;                                                                           // 放行脉冲预清 / Pass pulse preset
bError := FALSE;                                                                           // 故障标志预清（R45 配对） / Error preset
_iLen  := 0;                                                                               // 长度工作值预清 / Length working value preset

(* —— 段 2：组态闸（非法即锁存故障级） —— *)
IF _bCfgBad THEN
    _eCause := E_DL_FrcCause.eCfgIllegal;                                                  // 归因：组态非法 / Cause: illegal configuration
    _bFault := TRUE;                                                                       // 锁存 / Latch
    _eState := E_DL_FrcState.eFault;                                                       // 入故障相 / Enter fault phase
END_IF

(* —— 段 3：迁出链（bReset 上升沿：清双锁存，R228B） —— *)
IF rtReset.Q THEN
    _bFault := FALSE;                                                                      // 清故障锁存 / Clear fault latch
    _bFail  := FALSE;                                                                      // 清校验失败锁存 / Clear check-failure latch
    _eCause := E_DL_FrcCause.eNone;                                                        // 清成因 / Clear cause
    _eState := E_DL_FrcState.eIdle;                                                        // 回待机相 / Back to idle
END_IF

(* —— 段 4：相迁移（校验链；等待相三出口：读码沿 ∨ 超时 ∨ 启动撤销） —— *)
IF (NOT _bFault) AND (NOT _bCfgBad) THEN
    CASE _eState OF

    E_DL_FrcState.eIdle:
        IF rtStart.Q THEN
            _eState := E_DL_FrcState.eWait;                                                // 启动沿进等读码相 / Enter the wait phase
        END_IF

    E_DL_FrcState.eWait:
        IF rtRead.Q THEN
            (* —— 四段校验链（首因不覆盖：命中即锁存并停判） —— *)
            _iLen := LEN(sFoupId);                                                         // 取身份码长度 / Identity length
            IF _iLen = 0 THEN
                _bFail  := TRUE;                                                           // 失败锁存 / Latch the failure
                _eCause := E_DL_FrcCause.eIdEmpty;                                         // 首因：身份码空 / First cause: empty identity
            ELSIF (_iLen < UINT_TO_INT(uIdMinLen)) OR (_iLen > UINT_TO_INT(uIdMaxLen)) THEN
                _bFail  := TRUE;                                                           // 失败锁存 / Latch the failure
                _eCause := E_DL_FrcCause.eIdFormat;                                        // 首因：长度越域 / First cause: length out of range
            ELSIF LEN(sRecipeId) = 0 THEN
                _bFail  := TRUE;                                                           // 失败锁存 / Latch the failure
                _eCause := E_DL_FrcCause.eRecipeEmpty;                                     // 首因：在机配方空 / First cause: empty recipe
            ELSIF sRecipeId = sExpectedRecipe THEN
                _bPass  := TRUE;                                                           // 四段全过：放行脉冲（内部位） / All four checks passed
            ELSE
                _bFail  := TRUE;                                                           // 失败锁存 / Latch the failure
                _eCause := E_DL_FrcCause.eRecipeMismatch;                                  // 首因：配方不一致 / First cause: recipe mismatch
            END_IF

            IF _bFail THEN
                _bFault := TRUE;                                                           // 故障锁存 / Latch the fault
                _eState := E_DL_FrcState.eFault;                                           // 入故障相 / Enter fault phase
            ELSE
                _eState := E_DL_FrcState.eIdle;                                            // 放行后回待机相 / Back to idle after the pass
            END_IF
        ELSIF tonRead.Q THEN
            _bFail  := TRUE;                                                               // 读码超时：失败锁存 / Read timeout: latch the failure
            _eCause := E_DL_FrcCause.eReadTimeout;                                         // 首因：读码超时 / First cause: read timeout
            _bFault := TRUE;                                                               // 故障锁存 / Latch the fault
            _eState := E_DL_FrcState.eFault;                                               // 入故障相 / Enter fault phase
        ELSIF NOT bStartCheck THEN
            _eState := E_DL_FrcState.eIdle;                                                // 启动撤销：进相前置消失，回待机（出口 3，R129） / Start withdrawn, back to idle
        END_IF

    E_DL_FrcState.eFault:
        ;                                                                                  // 故障相：仅等复位沿 / Wait for the reset edge only

    ELSE
        _eCause := E_DL_FrcCause.ePhaseBad;                                                // 归因：非法相位 / Cause: illegal phase
        _bFault := TRUE;                                                                   // 锁存 / Latch
        _eState := E_DL_FrcState.eFault;                                                   // 强拉故障相 / Force fault phase

    END_CASE
END_IF

(* —— 段 5：出口单点映射（名实双出口，R191） —— *)
bPass        := _bPass;                                                                    // 放行脉冲出口 / Pass pulse outlet
bCheckFailed := _bFail;                                                                     // 校验失败出口 / Check-failure outlet
bWaiting     := (_eState = E_DL_FrcState.eWait);                                            // 等读码中出口 / Waiting outlet
eState       := _eState;                                                                    // 相出口 / Phase outlet
eCause       := _eCause;                                                                    // 成因出口 / Cause outlet
bError       := _bFault;                                                                    // 故障标志 / Error flag

END_FUNCTION_BLOCK

(* ---- FB_DL_FramingPressSeq.st ---- *)
(*
  FB_DL_FramingPressSeq  —  装框机压装顺控（涂胶-组框-压合节拍） / Framing press sequence: glue, frame, press cycle
  分类 Category : DL_Process
  版本 Version  : 1.0.0
  来源 Source   : t2-2-lbp — 层压/装框工艺族深化
  溯源 Origin   : clean-room 实现，未复制任何源码行
  功能 Function : 1) 四相顺控：eGlue（涂胶，等 bGlueDone 反馈）→ eFrame（组框定位，
                  等 bFrameDone 反馈）→ ePress（压合，合力窗判据）→ eDone → 回 eIdle；
                  2) 每相独立超时 TON（单相独占，R228-A），任一相超时 → 0374 锁存
                  （相推进超时同因族归并声明于码表）；压合相合力超上限当拍检出
                  → 0375 过载锁存（R146 方向独立：超上限走 0375，未达标走 0374）；
                  3) 信息级三码：序列启动 / 合力入窗 / 序列完成（单拍沿）；
                  4) 配比约束：tPressTo > tFrameTo > tGlueTo（压合节拍最长，
                  头注释按 R100 声明同拍三窗配比）；
                  5) 解除式全当拍量（R240 落地），逐 BOOL 标注见段 4。
  边界 Boundary : ① 组态闸：fForceMax <= fForceMin、任一超时 <= 0、或配比违反
                  （tPressTo <= tFrameTo 或 tFrameTo <= tGlueTo）→ 0373 锁存，
                  顺控全部停发，ELSE 兜底归并 0373（码表声明）；
                  ② 合力非有限 → 并入 0375 防御兜底（归并声明）；
                  ③ 相迁出仅由反馈当拍量承载，无锁存量自指；
                  ④ 无 GVL 依赖：纯引脚输入输出，无外部变量引用，无物理 IO 地址。
  依赖 Depends  : Standard.library（TON / R_TRIG）
  码表 Error codes（Process 段 0005，窗口 0373~0375 / 049B~049D）:
    16#0005_0373 故障级：组态非法（力窗颠倒/超时域/配比违反）或相位落 ELSE 兜底（归并声明），锁存至 bReset
    16#0005_0374 故障级：相推进超时（涂胶/组框/压合任一相独立计时到时，同因族归并声明），锁存至 bReset
    16#0005_0375 故障级：压合力过载超上限或合力非有限（防御兜底归并声明），锁存至 bReset
    16#0005_049B 信息级：压装序列启动沿（进 eGlue）
    16#0005_049C 信息级：压合力入窗沿（ePress 相）
    16#0005_049D 信息级：压装序列完成沿（进 eDone）
  修订历史 Revision :
    2026-11-19  v1.0.0  R42 首版（批次 1 · 序号 2）
*)

TYPE E_DL_FpsState :
(
    eIdle   := 0,    // 空闲：等启动沿 / Idle, waiting start edge
    eGlue   := 10,   // 涂胶：等涂胶完成反馈 / Glue, waiting glue-done feedback
    eFrame  := 20,   // 组框：等定位完成反馈 / Frame, waiting frame-done feedback
    ePress  := 30,   // 压合：合力窗判据 / Press, force band verdict
    eDone   := 40,   // 完成：序列落定 / Done
    eFault  := 90    // 故障：超时或过载锁定 / Fault, latched
);
END_TYPE

FUNCTION_BLOCK FB_DL_FramingPressSeq
VAR_INPUT
    bStart       : BOOL := FALSE;     // 启动指令，上升沿启动序列 [-] / Start command, rising edge
    bGlueDone    : BOOL := FALSE;     // 涂胶完成反馈（当拍量）[-] / Glue-done feedback
    bFrameDone   : BOOL := FALSE;     // 组框定位完成反馈（当拍量）[-] / Frame-done feedback
    fForceKgf    : REAL := 0.0;       // 压合合力反馈 [kgf]，调用方注入 / Press force feedback
    fForceMin    : REAL := 500.0;     // 合力窗下限 [kgf]，域 > 0 / Force band lower limit
    fForceMax    : REAL := 1200.0;    // 合力窗上限 [kgf]，必须 > fForceMin / Force band upper limit
    tGlueTo      : TIME := T#10S;     // 涂胶相超时 [ms]，域 > 0，配比最短 / Glue-phase timeout
    tFrameTo     : TIME := T#15S;     // 组框相超时 [ms]，域 > tGlueTo / Frame-phase timeout
    tPressTo     : TIME := T#20S;     // 压合相超时 [ms]，域 > tFrameTo / Press-phase timeout
    bReset       : BOOL := FALSE;     // 复位，上升沿清故障锁存 / Reset edge clears fault latch
END_VAR
VAR_OUTPUT
    eState       : E_DL_FpsState;     // 状态出口，段尾单点映射 / State outlet
    bRunning     : BOOL;              // 序列进行中标志（工艺相电平）[-] / Sequence running flag
    bDone        : BOOL;              // 序列完成标志（eDone 相电平）[-] / Sequence done flag
    bForceInBand : BOOL;              // 合力入窗实时镜像 [-] / Force-in-band mirror
    bError       : BOOL;              // 故障锁存标志 / Fault latch flag
    nErrId       : UDINT;             // 事件码，0 = 无事件 / Event code
END_VAR
VAR
    tonGlueTo    : TON;               // 涂胶相超时（单相独占），无条件刷新 / Glue-phase timeout
    tonFrameTo   : TON;               // 组框相超时（单相独占），无条件刷新 / Frame-phase timeout
    tonPressTo   : TON;               // 压合相超时（单相独占），无条件刷新 / Press-phase timeout
    rtStart      : R_TRIG;            // 启动沿实例，无条件刷新 / Start edge instance
    rtReset      : R_TRIG;            // 复位沿实例，无条件刷新 / Reset edge instance
    _eState      : E_DL_FpsState := E_DL_FpsState.eIdle;  // 内部相位（CASE 唯一写入目标）/ Internal phase
    _bForceOk    : BOOL;              // 合力入窗当拍量 [-] / Force-in-band current-scan flag
    _bOver       : BOOL;              // 合力超上限当拍量 [-] / Force-over-limit current-scan flag
    _bNonFin     : BOOL;              // 合力非有限当拍量 [-] / Non-finite force current-scan flag
    _bFault      : BOOL;              // 故障锁存位（锁存量）/ Latched fault bit
    _uFault      : UDINT;             // 故障码锁存（锁存量）/ Latched fault code
    _uInfo       : UDINT;             // 信息码，每拍重算 / Transient info code
END_VAR

(* —— 段 0：定时器与沿实例无条件周期刷新（禁置于 IF/CASE 内） —— *)
_bForceOk := (fForceKgf >= fForceMin) AND (fForceKgf <= fForceMax);  // 合力入窗（当拍量）
_bOver   := fForceKgf > fForceMax;                                   // 过载方向独立检出（R146）
_bNonFin := (fForceKgf <> fForceKgf)
         OR ((fForceKgf - fForceKgf) <> (fForceKgf - fForceKgf));    // 非有限防御（NaN 自反 + 差值自减）
rtStart(CLK := bStart);                                              // 启动沿（每拍必调）
rtReset(CLK := bReset);                                              // 复位沿（每拍必调）
tonGlueTo(IN := (_eState = E_DL_FpsState.eGlue), PT := tGlueTo);     // 涂胶相超时（单相独占）
tonFrameTo(IN := (_eState = E_DL_FpsState.eFrame), PT := tFrameTo);  // 组框相超时（单相独占）
tonPressTo(IN := (_eState = E_DL_FpsState.ePress), PT := tPressTo);  // 压合相超时（单相独占）

(* —— 段 1：单拍量预清零（锁存量 _bFault/_uFault 不入清单，禁同拍抹除） —— *)
_uInfo := 16#0000_0000;             // 信息码每拍重算
bRunning := FALSE;                  // 进行中标志缺省 FALSE
bDone := FALSE;                     // 完成标志缺省 FALSE
bForceInBand := FALSE;              // 入窗镜像缺省 FALSE
nErrId := 16#0000_0000;             // 事件码缺省无事件

(* —— 段 2：复位沿 + 组态域闸（当拍量判据，含 R100 配比约束） —— *)
IF rtReset.Q THEN                   // rtReset.Q = 当拍量
    _bFault := FALSE;               // 清故障锁存位
    _uFault := 16#0000_0000;        // 清故障锁存码
END_IF
IF (fForceMax <= fForceMin) OR (TIME_TO_DINT(tGlueTo) <= 0)
   OR (TIME_TO_DINT(tFrameTo) <= 0) OR (TIME_TO_DINT(tPressTo) <= 0)
   OR (tPressTo <= tFrameTo) OR (tFrameTo <= tGlueTo) THEN
    _uFault := 16#0005_0373;        // 故障级：组态非法（含配比违反）
    _bFault := TRUE;                // 故障标志与码位配对（R45）
END_IF

(* —— 段 3：相超时与过载锁存（判据当拍量/单相独占 TON） —— *)
IF (NOT _bFault) AND (tonGlueTo.Q OR tonFrameTo.Q OR tonPressTo.Q) THEN
    _uFault := 16#0005_0374;        // 故障级：相推进超时（同因族归并声明）
    _bFault := TRUE;
END_IF
IF (NOT _bFault) AND (_eState = E_DL_FpsState.ePress) AND (_bOver OR _bNonFin) THEN
    _uFault := 16#0005_0375;        // 故障级：压合力过载或非有限（防御兜底归并）
    _bFault := TRUE;
END_IF

(* —— 段 4：故障解除式（R240 落地，逐 BOOL 标注）：
     rtReset.Q = 当拍量；bStart = 当拍量；均不含锁存量（_bFault/_uFault），
     解除边真实可达（启动指令撤销后复位沿可到达）。 —— *)
IF rtReset.Q AND (NOT bStart) THEN
    _bFault := FALSE;               // 清故障锁存位（锁存量，仅此当拍量解除沿可清）
    _uFault := 16#0000_0000;        // 清故障锁存码（锁存量，仅本当拍量解除沿可清）
    IF _eState = E_DL_FpsState.eFault THEN
        _eState := E_DL_FpsState.eIdle;     // 故障相迁出：回空闲
    END_IF
END_IF

(* —— 段 5：相位机（CASE 全覆盖 + ELSE 兜底） —— *)
CASE _eState OF

E_DL_FpsState.eIdle:
    IF rtStart.Q AND (NOT _bFault) THEN
        _uInfo := 16#0005_049B;             // 信息级：序列启动沿
        _eState := E_DL_FpsState.eGlue;     // 进涂胶相
    END_IF

E_DL_FpsState.eGlue:
    bRunning := TRUE;                       // 进行中标志（相电平）
    IF bGlueDone THEN
        _eState := E_DL_FpsState.eFrame;    // 涂胶完成：进组框相
    END_IF
    (* 超时迁出在段 3 承载 *)

E_DL_FpsState.eFrame:
    bRunning := TRUE;                       // 进行中标志（相电平）
    IF bFrameDone THEN
        _eState := E_DL_FpsState.ePress;    // 定位完成：进压合相
    END_IF

E_DL_FpsState.ePress:
    bRunning := TRUE;                       // 进行中标志（相电平）
    bForceInBand := _bForceOk;              // 入窗镜像（相电平）
    IF _bForceOk THEN
        _uInfo := 16#0005_049C;             // 信息级：合力入窗沿
        _eState := E_DL_FpsState.eDone;     // 判据达成：进完成相
    END_IF
    (* 过载迁出在段 3 承载 *)

E_DL_FpsState.eDone:
    bDone := TRUE;                          // 完成标志（相电平）
    _uInfo := 16#0005_049D;                 // 信息级：序列完成（相电平重发，信息级允许）
    IF NOT bStart THEN                      // 启动指令撤销：回空闲
        _eState := E_DL_FpsState.eIdle;
    END_IF

E_DL_FpsState.eFault:
    ;                                       // 故障相：等复位沿（段 4 承载迁出）

ELSE
    _uFault := 16#0005_0373;                // 故障级：非法相位兜底（归并组态码，码表声明）
    _bFault := TRUE;
    _eState := E_DL_FpsState.eFault;        // 强制回故障相

END_CASE

(* —— 段 6：出口单点映射（名实同源；锁存码回放，禁同拍抹除） —— *)
IF _bFault THEN
    nErrId := _uFault;              // 故障锁存码回放
    bRunning := FALSE;              // 故障相进行中出口强制 FALSE（安全侧）
    bDone := FALSE;                 // 故障相完成出口强制 FALSE（安全侧）
    bForceInBand := FALSE;          // 故障相入窗镜像强制 FALSE（安全侧）
ELSE
    nErrId := _uInfo;               // 信息码
END_IF
bError := _bFault;                  // 故障标志与锁存位同源
eState := _eState;                  // 状态出口单点映射

END_FUNCTION_BLOCK

(* ---- FB_DL_FreezeStatGuard.st ---- *)
(*
  Component : FB_DL_FreezeStatGuard
  Category  : DL_Process
  Type      : FB
  Version   : 1.0.0
  CodeSeg   : 16#06_0_38
  Summary   : 表冷器防冻保护与低温联锁：低温门限持续判定 + 预热阀比例调节 + 冻结告警锁存。
              Coil freeze protection: sustained low-temp gate plus proportional preheat valve and latched freeze alarm.
  溯源声明  : 道莅自研 clean-room
  边界安全  : 温度非有限（NaN 自反 + Inf 上限）拦截；低温需持续 tFrostMs（TON 防单拍毛刺误报）；
              预热阀输出钳 0..100 ％；冻结告警锁存且解除路径可达（温度恢复 + 复位沿）；
              TON/R_TRIG 每拍无条件刷新（段 0）；全浮点比较带 fEps 容差。
  复用      : 无
*)

FUNCTION_BLOCK FB_DL_FreezeStatGuard
VAR_INPUT
    bRun       : BOOL;                  (* 保护使能 · Enable *)
    fAirTC     : LREAL;                 (* 表冷器后风温 [degC] · Coil downstream air temperature *)
    fFrostThC  : LREAL := 2.0;          (* 低温门限 [degC] · Low temperature threshold *)
    fGainPctK  : LREAL := 25.0;         (* 预热阀比例增益 [％/K] · Preheat proportional gain *)
    tFrostMs   : TIME  := T#10000MS;    (* 低温持续窗 [ms] · Sustained low-temp window *)
    bReset     : BOOL;                  (* 告警复位指令 [事件]，沿触发 · Alarm reset command *)
    fEps       : LREAL := 1.0E-6;       (* 浮点判零容差 [实数域] · Floating zero tolerance *)
END_VAR
VAR_OUTPUT
    fPreheatPct: LREAL;                 (* 预热阀开度输出 [％] · Preheat valve output *)
    bPreheat   : BOOL;                  (* 预热激活标志 · Preheat active flag *)
    bFrostWarn : BOOL;                  (* 低温持续告警（非锁存）· Sustained frost warning *)
    bFreezeAlm : BOOL;                  (* 冻结告警锁存 · Latched freeze alarm *)
    bError     : BOOL;                  (* 故障标志，与故障码配对 · Fault flag paired with codes *)
    uErrorId   : UDINT;                 (* 事件码 16#0000_0038，0 无事件 · Event code *)
END_VAR
VAR
    _eState  : (eStWatch := 0, eStFrozen := 1);     (* 内部状态机 / Internal state machine *)
    uCode    : WORD;    (* 码位暂存，每拍重算 [码] · Code staging *)
    tonFrost : TON;     (* 低温持续计时 [ms]，每拍无条件刷新 · Frost duration timer *)
    rTrigRst : R_TRIG;  (* 复位沿检测 · Reset edge detection *)
    bSigOk   : BOOL;    (* 输入有效标志 · Input validity flag *)
    bLowNow  : BOOL;    (* 本拍低温判定 / This-scan low-temp verdict *)
    fSubK    : LREAL;   (* 过冷深度 [K] · Sub-cooling depth *)
    nCycles  : UDINT;   (* 有效监视拍计数 [拍]，防回卷 · Monitor scan count *)
END_VAR
VAR CONSTANT
    DL_FSG_WRAP : UDINT := 4294967290;  (* 计数防回卷余量 [拍] · Counter wrap guard *)
    DL_FSG_PCTMAX: LREAL := 100.0;      (* 阀开度上限 [％] · Valve output cap *)
END_VAR

(* === 段 0 · 实例刷新（每拍无条件，红线 7）=== *)
tonFrost(IN := bRun AND bSigOk AND (NOT bFreezeAlm), PT := tFrostMs);   (* 低温持续计时 / Frost timing *)
rTrigRst(CLK := bReset);                        (* 复位沿检测 / Reset edge *)

(* === 段 1 · 输入校验与量程闸 === *)
uCode := 16#0000;                       // 每拍清码（可达清零基线）/ Clear codes each scan
bSigOk := (fAirTC = fAirTC) AND (ABS(fAirTC) < 1.0E308)             // 非有限拦截 / Non-finite guard
          AND (fFrostThC = fFrostThC) AND (fGainPctK >= 0.0)         // 门限非有限 + 增益非负闸 / Threshold and gain gates
          AND (tFrostMs > T#0MS);                                    (* 持续窗正域闸 / Duration window gate *)
IF NOT bSigOk THEN
    uCode := 16#0038;                   // 故障级：域外，保护冻结于安全输出 / Fault: domain invalid
END_IF

(* === 段 2 · 主逻辑：低温判定与冻结告警状态机 === *)
IF bSigOk THEN
    bLowNow := (fAirTC < fFrostThC);    (* 本拍低温判定（单比较非容差问题）/ Low-temp verdict *)
    fSubK := fFrostThC - fAirTC;        (* 过冷深度 [K] / Sub-cooling depth *)
    IF fSubK < 0.0 THEN
        fSubK := 0.0;                   (* 深度钳非负 / Clamp non-negative *)
    END_IF
    CASE _eState OF
        eStWatch:                       (* 监视相：低温持续到点转冻结 / Watch: escalate on sustained frost *)
            IF tonFrost.Q THEN
                _eState := eStFrozen;   (* 拍 N 窗满，拍 N+1 转冻结相 / To frozen next scan *)
            END_IF
        eStFrozen:                      (* 冻结相：告警锁存 / Frozen: alarm latched *)
            (* 解除路径：温度恢复 + 复位沿（可达）/ Clear: recovery plus reset edge *)
            IF rTrigRst.Q AND (NOT bLowNow) THEN
                _eState := eStWatch;    (* 拍 N+1 回监视相 / Back to watch *)
            END_IF
    ELSE
        _eState := eStWatch;            (* ELSE 兜底回监视相 / ELSE fallback to watch *)
        uCode := 16#0038;               (* 状态越界报码 / Code on illegal state *)
    END_CASE
    bFreezeAlm := (_eState = eStFrozen);        (* 冻结告警回放 / Latched alarm replay *)
    bFrostWarn := tonFrost.Q;           (* 低温持续告警（非锁存自清）/ Non-latched warning *)
    (* 预热阀比例调节：过冷深度 × 增益，冻结相全开 / Proportional preheat, full open when frozen *)
    IF bFreezeAlm THEN
        fPreheatPct := DL_FSG_PCTMAX;   (* 冻结全开预热 / Full open when frozen *)
    ELSIF bLowNow THEN
        fPreheatPct := fSubK * fGainPctK;   (* 比例调节 [％] / Proportional output *)
        IF fPreheatPct > DL_FSG_PCTMAX THEN
            fPreheatPct := DL_FSG_PCTMAX;   (* 钳上限 / Cap high *)
        END_IF
    ELSE
        fPreheatPct := 0.0;             (* 正温关阀 / Close on normal temperature *)
    END_IF
END_IF

(* === 段 3 · 输出映射与故障码 === *)
IF NOT bRun THEN
    bFreezeAlm := FALSE;                (* 撤使能告警释放（可达清零路径）/ Clear on disable *)
    _eState := eStWatch;                (* 回监视相 / Back to watch *)
    fPreheatPct := 0.0;                 (* 阀关安全位 / Safe valve close *)
END_IF
bPreheat := (fPreheatPct > fEps);       (* 预热激活标志 / Preheat active flag *)
IF bSigOk THEN
    IF nCycles < DL_FSG_WRAP THEN
        nCycles := nCycles + 1;         (* 有效监视计数 / Count monitor scans *)
    END_IF
END_IF
bError := bFreezeAlm OR (uCode <> 16#0000);     (* 故障标志 / Fault flag *)
IF bFreezeAlm THEN
    uErrorId := WORD_TO_UDINT(16#0038); (* 码位 16#0000_0038 冻结告警 / Freeze alarm code *)
ELSE
    uErrorId := WORD_TO_UDINT(uCode);   (* 域外码或零 / Domain code or zero *)
END_IF
END_FUNCTION_BLOCK

(* ---- FB_DL_FurnaceDoorInterlockSeq.st ---- *)
(*
  Name: FB_DL_FurnaceDoorInterlockSeq
  Category: DL_Process
  Version: 1.0.0
  Round: R89 / 2026-11-25
  开源溯源：clean-room 自研（族 锻造加热退火，ST 开源生态实测 0 命中，无外部代码引入）
  功能：炉门与气氛/温度联锁开关顺序：开门前必须先断气氛、并降到安全温度以下、且炉内无正压。
  边界条件：① 三浮点入参全部过非有限闸；配置越域即锁故障（101）；
            ② 顺序强制：气氛未断不降温等待、温度未降到「安全温度 − 20 ℃」不给开门许可（带回差防抖）；
            ③ 正压（> 2.0 kPa）时禁止开门并锁故障（102），须泄压后重新申请；
            ④ 开门许可相内若温度回升或气氛复投，立即撤回许可并退回冷却等待相（安全侧优先）；
            ⑤ 故障解除唯一路径：故障相内 xOpenCmd 释放（R152），清锁存回 eIdle。
  状态机：eIdle / eAtmosCut / eCoolWait / eDoorPermit / eFault（CASE 含 ELSE 兜底）。
*)
TYPE E_DL_FdiState :
(
    eIdle      := 0,    (* 待机：等开门申请 / Idle, waiting for open request *)
    eAtmosCut  := 10,   (* 断气氛相：等气氛阀关闭反馈 / Atmos cut, waiting feedback *)
    eCoolWait  := 20,   (* 降温等待相：等温度降到安全值以下 / Cooling wait *)
    eDoorPermit := 30,  (* 开门许可相：允许开炉门 / Door permit *)
    eFault     := 90    (* 故障相：锁存待释放 / Fault latched, awaiting release *)
);
END_TYPE

FUNCTION_BLOCK FB_DL_FurnaceDoorInterlockSeq
VAR_INPUT
    xOpenCmd : BOOL;        (* 开门申请 [-] Door open request *)
    fTempC : REAL;          (* 炉内温度实测 [℃] Furnace temperature actual [degC] *)
    fTempSafeC : REAL;      (* 安全开门温度 [℃] Safe opening temperature [degC] *)
    xAtmosOn : BOOL;        (* 气氛投入反馈（TRUE = 已投） [-] Atmosphere on feedback *)
    fPressKPa : REAL;       (* 炉内压力（表压） [kPa] Furnace gauge pressure [kPa] *)
END_VAR
VAR_OUTPUT
    xDoorPermit : BOOL;     (* 开门许可 [-] Door permit *)
    xAtmosCutCmd : BOOL;    (* 断气氛指令（顺序期间保持） [-] Atmosphere cut command *)
    xFault : BOOL;          (* 故障锁存标志 [-] Fault latched *)
    nErrCode : INT;         (* 故障码 0/101 组态/102 正压超限/103 非法相 [-] Error code *)
END_VAR
VAR
    _eState : E_DL_FdiState := E_DL_FdiState.eIdle;  (* 内部相（CASE 唯一写入目标） [-] Internal phase *)
    _bFaultLatch : BOOL := FALSE;   (* 故障锁存位 [-] Fault latch *)
    _bReqFault : BOOL := FALSE;     (* 单拍故障请求（段 1 预清） [-] Fault request *)
    _bCfgBad : BOOL := FALSE;       (* 组态非法当拍量 [-] Configuration bad *)
    _bTempSafe : BOOL := FALSE;     (* 温度已降到安全值以下 [-] Temperature below safe value *)
    _bPressOk : BOOL := FALSE;      (* 炉内无正压 [-] No positive pressure *)
    _nErr : INT := 0;               (* 故障码锁存 [-] Latched error code *)
    _nReqErr : INT := 0;            (* 当拍请求码 [-] Requested error code *)
END_VAR
VAR CONSTANT
    DL_FDI_HYST : REAL := 20.0;     (* 安全温度回差 [℃] Safety temperature hysteresis [degC] *)
    DL_FDI_PMAX : REAL := 2.0;      (* 允许开门正压上限 [kPa] Allowed positive pressure [kPa] *)
    DL_FDI_TS_MIN : REAL := 20.0;   (* 安全温度下限 [℃] Safe temperature floor [degC] *)
    DL_FDI_TS_MAX : REAL := 200.0;  (* 安全温度上限 [℃] Safe temperature ceiling [degC] *)
    DL_FDI_T_MIN : REAL := -50.0;   (* 炉温下限 [℃] Furnace temperature floor [degC] *)
    DL_FDI_T_MAX : REAL := 1400.0;  (* 炉温上限 [℃] Furnace temperature ceiling [degC] *)
    DL_FDI_P_MIN : REAL := -5.0;    (* 压力量程下限 [kPa] Pressure floor [kPa] *)
    DL_FDI_P_MAX : REAL := 5.0;     (* 压力量程上限 [kPa] Pressure ceiling [kPa] *)
END_VAR
(* —— 段 0：非有限闸（NaN 自反 + Inf 差值自减）+ 组态域闸，三浮点入参全枚举（R272） —— *)
_bCfgBad := (fTempC <> fTempC) OR ((fTempC - fTempC) <> 0.0)
         OR (fTempSafeC <> fTempSafeC) OR ((fTempSafeC - fTempSafeC) <> 0.0)
         OR (fPressKPa <> fPressKPa) OR ((fPressKPa - fPressKPa) <> 0.0)
         OR (fTempC < DL_FDI_T_MIN) OR (fTempC > DL_FDI_T_MAX)
         OR (fTempSafeC < DL_FDI_TS_MIN) OR (fTempSafeC > DL_FDI_TS_MAX)
         OR (fPressKPa < DL_FDI_P_MIN) OR (fPressKPa > DL_FDI_P_MAX);
(* 两个判据量：温度须低于「安全温度 − 回差」；压力须不超过允许正压 *)
_bTempSafe := fTempC <= (fTempSafeC - DL_FDI_HYST);
_bPressOk := fPressKPa <= DL_FDI_PMAX;
(* —— 段 1：单拍量预清 + 组态故障请求 —— *)
_bReqFault := FALSE;
_nReqErr := 0;
IF _bCfgBad THEN
    _bReqFault := TRUE; _nReqErr := 101;        (* 组态非法 / Configuration bad *)
END_IF
(* —— 段 2：故障锁存解除（唯一路径 = 故障相内 xOpenCmd 释放，R152） —— *)
IF _bFaultLatch AND (NOT xOpenCmd) THEN
    _bFaultLatch := FALSE;                      (* 清锁存 / Clear latch *)
    _nErr := 0;                                 (* 清码 / Clear code *)
    _eState := E_DL_FdiState.eIdle;             (* 迁回待机 / Back to idle *)
END_IF
(* —— 段 3：主状态机（ENUM + CASE，ELSE 兜底） —— *)
CASE _eState OF
E_DL_FdiState.eIdle:
    IF xOpenCmd AND (NOT _bFaultLatch) THEN
        IF xAtmosOn THEN
            _eState := E_DL_FdiState.eAtmosCut; (* 已投气氛：先断气氛 / Atmosphere on, cut first *)
        ELSE
            _eState := E_DL_FdiState.eCoolWait; (* 未投气氛：直接降温等待 / No atmos, cool wait *)
        END_IF
    END_IF
E_DL_FdiState.eAtmosCut:
    IF NOT xAtmosOn THEN
        _eState := E_DL_FdiState.eCoolWait;     (* 气氛已断 → 降温等待 / Atmos off, cool wait *)
    END_IF
E_DL_FdiState.eCoolWait:
    IF (NOT xAtmosOn) AND _bTempSafe THEN
        IF _bPressOk THEN
            _eState := E_DL_FdiState.eDoorPermit;   (* 三项齐备 → 开门许可 / All ready, permit *)
        ELSE
            _bReqFault := TRUE; _nReqErr := 102;    (* 正压超限：禁止开门 / Positive pressure *)
        END_IF
    END_IF
E_DL_FdiState.eDoorPermit:
    IF NOT xOpenCmd THEN
        _eState := E_DL_FdiState.eIdle;         (* 申请撤销 → 待机 / Request withdrawn *)
    ELSIF xAtmosOn OR (NOT _bTempSafe) OR (NOT _bPressOk) THEN
        _eState := E_DL_FdiState.eCoolWait;     (* 前置失守 → 退回等待（安全侧优先） / Precondition lost *)
    END_IF
E_DL_FdiState.eFault:
    _bPressOk := fPressKPa <= DL_FDI_PMAX;      (* 故障相驻留：判据照算供追溯，不迁相 *)
ELSE
    _bReqFault := TRUE;                         (* 非法相兜底 / Illegal phase fallback *)
    _nReqErr := 103;
END_CASE
(* —— 段 4：故障请求统一落地（唯一锁存点 + 同步迁相，R187/R252） —— *)
IF _bReqFault AND (NOT _bFaultLatch) THEN
    _bFaultLatch := TRUE;                       (* 锁存 / Latch *)
    _nErr := _nReqErr;                          (* 码锁存回放 / Latched code *)
    _eState := E_DL_FdiState.eFault;            (* 同步迁相 / Migrate to fault *)
END_IF
(* —— 段 5：统一出口（各出口单点赋值） —— *)
xDoorPermit := (_eState = E_DL_FdiState.eDoorPermit) AND (NOT _bFaultLatch);
xAtmosCutCmd := (_eState = E_DL_FdiState.eAtmosCut) OR (_eState = E_DL_FdiState.eCoolWait)
             OR (_eState = E_DL_FdiState.eDoorPermit);
xFault := _bFaultLatch;
nErrCode := _nErr;
END_FUNCTION_BLOCK

(* ---- FB_DL_FurnaceZoneHeatSeq.st ---- *)
(*
  Name: FB_DL_FurnaceZoneHeatSeq
  Category: DL_Process
  Version: 1.0.0
  Round: R89 / 2026-11-25
  开源溯源：clean-room 自研（族 锻造加热退火，ST 开源生态实测 0 命中，无外部代码引入）
  功能：多区加热炉分区升温监视与顺序校核：每区独立稳态判定，低温区未到位而高温区先到即判顺序违例。
  边界条件：① 八浮点入参（四区实测 + 四区设定）与公差、稳态窗全部过非有限闸；
            ② 每区独立 TON（tonZ1~tonZ4），PT 均取 tSettleS，禁跨区共用（R100 无同拍双窗）；
            ③ 顺序判据：区 i 已进带而存在设定更低（低 1 ℃ 以上）的区 j 尚未进带 → 违例 → 锁故障；
            ④ 故障解除唯一路径：故障相内 xStart 释放（R152），清锁存回 eIdle。
  状态机：eIdle / eHeat / eAllReady / eFault（CASE 含 ELSE 兜底）。
*)
TYPE E_DL_FzsState :
(
    eIdle     := 0,     (* 待机：等启动沿 / Idle, waiting for start edge *)
    eHeat     := 10,    (* 升温监视相：逐区稳态计时与顺序校核 / Heat monitoring *)
    eAllReady := 20,    (* 全区到位相：保持至启动释放 / All zones ready, holds *)
    eFault    := 90     (* 故障相：锁存待释放 / Fault latched, awaiting release *)
);
END_TYPE

FUNCTION_BLOCK FB_DL_FurnaceZoneHeatSeq
VAR_INPUT
    xStart : BOOL;                          (* 启动命令（上升沿起序） [-] Start command, rising edge *)
    anZoneTempC : ARRAY[1..4] OF REAL;      (* 四区实测温度 [℃] Zone temperatures [degC] *)
    fZoneSpC : ARRAY[1..4] OF REAL;         (* 四区设定温度 [℃] Zone setpoints [degC] *)
    fDevTolC : REAL;                        (* 稳态带半宽 [℃] Steady band half-width [degC] *)
    tSettleS : TIME;                        (* 单区稳态窗 [ms] Per-zone settling window [ms] *)
END_VAR
VAR_OUTPUT
    eState : E_DL_FzsState;                 (* 当前相 [-] Present phase *)
    nZoneReady : INT;                       (* 已稳态到位的区数（0~4） [区] Ready zone count *)
    xAllReady : BOOL;                       (* 四区全部到位 [-] All zones ready *)
    xFault : BOOL;                          (* 故障锁存标志 [-] Fault latched *)
END_VAR
VAR
    _eState : E_DL_FzsState := E_DL_FzsState.eIdle;  (* 内部相（CASE 唯一写入目标） [-] Internal phase *)
    _abBand : ARRAY[1..4] OF BOOL;          (* 各区在稳态带内 [-] Zone in steady band *)
    _abSettled : ARRAY[1..4] OF BOOL;       (* 各区稳态窗已满 [-] Zone settled *)
    _bFaultLatch : BOOL := FALSE;           (* 故障锁存位 [-] Fault latch *)
    _bCfgBad : BOOL := FALSE;               (* 组态非法当拍量 [-] Configuration bad *)
    _bOrderViol : BOOL := FALSE;            (* 升温顺序违例 [-] Heating order violation *)
    _bAllReady : BOOL := FALSE;             (* 全区到位当拍量 [-] All ready this scan *)
    _nReady : INT := 0;                     (* 到位区计数 [区] Ready count *)
    _nI : INT := 1;                         (* 区遍历索引（外层） [-] Outer loop index *)
    _nJ : INT := 1;                         (* 区遍历索引（内层） [-] Inner loop index *)
    tonZ1 : TON;                            (* 一区稳态窗（段 0 无条件调用） / Zone 1 window *)
    tonZ2 : TON;                            (* 二区稳态窗（段 0 无条件调用） / Zone 2 window *)
    tonZ3 : TON;                            (* 三区稳态窗（段 0 无条件调用） / Zone 3 window *)
    tonZ4 : TON;                            (* 四区稳态窗（段 0 无条件调用） / Zone 4 window *)
    rtStart : R_TRIG;                       (* 启动沿（段 0 无条件调用） / Start edge *)
END_VAR
VAR CONSTANT
    DL_FZS_TOL_MIN : REAL := 0.5;       (* 稳态带半宽下限 [℃] Band floor [degC] *)
    DL_FZS_TOL_MAX : REAL := 50.0;      (* 稳态带半宽上限 [℃] Band ceiling [degC] *)
    DL_FZS_SP_MIN : REAL := 50.0;       (* 设定温度下限 [℃] Setpoint floor [degC] *)
    DL_FZS_SP_MAX : REAL := 1350.0;     (* 设定温度上限 [℃] Setpoint ceiling [degC] *)
    DL_FZS_ORD : REAL := 1.0;           (* 顺序比较死区（设定差大于此值才判前后） [℃] Order deadband [degC] *)
    DL_FZS_ZNUM : INT := 4;             (* 分区总数 [-] Zone count *)
END_VAR
(* —— 段 0：沿与四区稳态 TON 无条件周期刷新（R7），IN 由带内判据与相位共同派生 —— *)
rtStart(CLK := xStart);                                                     (* 启动沿 / Start edge *)
(* 带内判据：逐区算（NaN 与非有限在下面组态闸统一拦截，此处比较对 NaN 恒假即不进带） *)
FOR _nI := 1 TO DL_FZS_ZNUM DO
    _abBand[_nI] := (anZoneTempC[_nI] = anZoneTempC[_nI]) AND (ABS(anZoneTempC[_nI] - fZoneSpC[_nI]) <= fDevTolC);
END_FOR
tonZ1(IN := _abBand[1] AND (_eState = E_DL_FzsState.eHeat), PT := tSettleS);   (* 一区稳态窗 / Zone 1 *)
tonZ2(IN := _abBand[2] AND (_eState = E_DL_FzsState.eHeat), PT := tSettleS);   (* 二区稳态窗 / Zone 2 *)
tonZ3(IN := _abBand[3] AND (_eState = E_DL_FzsState.eHeat), PT := tSettleS);   (* 三区稳态窗 / Zone 3 *)
tonZ4(IN := _abBand[4] AND (_eState = E_DL_FzsState.eHeat), PT := tSettleS);   (* 四区稳态窗 / Zone 4 *)
_abSettled[1] := tonZ1.Q;                   (* 一区到位 / Zone 1 settled *)
_abSettled[2] := tonZ2.Q;                   (* 二区到位 / Zone 2 settled *)
_abSettled[3] := tonZ3.Q;                   (* 三区到位 / Zone 3 settled *)
_abSettled[4] := tonZ4.Q;                   (* 四区到位 / Zone 4 settled *)
(* 非有限闸 + 组态域闸：公差、稳态窗与八区温度量全枚举（R272） *)
_bCfgBad := (fDevTolC <> fDevTolC) OR ((fDevTolC - fDevTolC) <> 0.0)
         OR (fDevTolC < DL_FZS_TOL_MIN) OR (fDevTolC > DL_FZS_TOL_MAX)
         OR (tSettleS <= T#0S);
FOR _nI := 1 TO DL_FZS_ZNUM DO
    IF (anZoneTempC[_nI] <> anZoneTempC[_nI]) OR ((anZoneTempC[_nI] - anZoneTempC[_nI]) <> 0.0)
       OR (fZoneSpC[_nI] <> fZoneSpC[_nI]) OR ((fZoneSpC[_nI] - fZoneSpC[_nI]) <> 0.0)
       OR (fZoneSpC[_nI] < DL_FZS_SP_MIN) OR (fZoneSpC[_nI] > DL_FZS_SP_MAX) THEN
        _bCfgBad := TRUE;
    END_IF
END_FOR
(* 顺序校核：区 i 已进带，而存在设定更低（低 DL_FZS_ORD 以上）的区 j 尚未进带 → 违例 *)
_bOrderViol := FALSE;
FOR _nI := 1 TO DL_FZS_ZNUM DO
    IF _abBand[_nI] THEN
        FOR _nJ := 1 TO DL_FZS_ZNUM DO
            IF (fZoneSpC[_nJ] < (fZoneSpC[_nI] - DL_FZS_ORD)) AND (NOT _abBand[_nJ]) THEN
                _bOrderViol := TRUE;
            END_IF
        END_FOR
    END_IF
END_FOR
(* 到位计数：稳态窗满即计入 *)
_nReady := 0;
FOR _nI := 1 TO DL_FZS_ZNUM DO
    IF _abSettled[_nI] THEN
        _nReady := _nReady + 1;
    END_IF
END_FOR
_bAllReady := (_nReady = DL_FZS_ZNUM);
(* —— 段 1：单拍量预清 + 组态/顺序故障请求 —— *)
IF _bCfgBad OR _bOrderViol THEN
    _bFaultLatch := TRUE;                   (* 锁存 / Latch *)
END_IF
(* —— 段 2：故障锁存解除（唯一路径 = 故障相内 xStart 释放，R152） —— *)
IF _bFaultLatch AND (NOT xStart) THEN
    _bFaultLatch := FALSE;                  (* 清锁存 / Clear latch *)
    _eState := E_DL_FzsState.eIdle;         (* 迁回待机 / Back to idle *)
END_IF
(* —— 段 3：主状态机（ENUM + CASE，ELSE 兜底） —— *)
CASE _eState OF
E_DL_FzsState.eIdle:
    IF rtStart.Q AND (NOT _bFaultLatch) THEN
        _eState := E_DL_FzsState.eHeat;     (* 起序 → 升温监视 / Start, heat monitoring *)
    END_IF
E_DL_FzsState.eHeat:
    IF _bFaultLatch THEN
        _eState := E_DL_FzsState.eFault;    (* 违例/组态坏 → 故障 / Violation, to fault *)
    ELSIF _bAllReady THEN
        _eState := E_DL_FzsState.eAllReady; (* 全区到位 → 到位相 / All ready *)
    END_IF
E_DL_FzsState.eAllReady:
    IF NOT xStart THEN
        _eState := E_DL_FzsState.eIdle;     (* 启动释放 → 待机 / Start released, idle *)
    END_IF
E_DL_FzsState.eFault:
    _bAllReady := (_nReady = DL_FZS_ZNUM);  (* 故障相驻留：到位判据照算供追溯，不迁相 *)
ELSE
    _bFaultLatch := TRUE;                   (* 非法相兜底 / Illegal phase fallback *)
    _eState := E_DL_FzsState.eFault;
END_CASE
(* —— 段 4：统一出口（各出口单点赋值） —— *)
eState := _eState;
nZoneReady := _nReady;
xAllReady := _bAllReady AND (NOT _bFaultLatch);
xFault := _bFaultLatch;
END_FUNCTION_BLOCK

(* ---- FB_DL_GlassFeederAccum.st ---- *)
(*
  FB_DL_GlassFeederAccum  —  玻璃上料输送积放（多区级联积放协调） / Glass feeder multi-zone accumulation and cascade release coordinator
  分类 Category : DL_Process
  版本 Version  : 1.0.0
  来源 Source   : t2-2-lbp — 玻璃输送/积放族深化
  溯源 Origin   : clean-room 实现，未复制任何源码行
  功能 Function : 1) 四区级联积放：eIdle（积放保持，挡板全抬起）→ eRel（放行序列：
                  自下游区 0 起逐区落挡板放行、等区光电放空、抬板进下一区）
                  → 全区放空回 eIdle；
                  2) 释放相单区超时 tZoneTo → 037D 锁存（R233 单相独占分实例）；
                  3) 积放相背压监视：非释放相全部区占满且输送运行持续 tAccumTo
                  → 037E 满载滞留锁存（归因独立于释放超时）；
                  4) 信息级三码：积放激活 / 区释放沿 / 全区放行完成；
                  5) 解除式全当拍量（R240 落地），逐 BOOL 标注见段 4。
  边界 Boundary : ① 组态闸：任一时间 <= 0 → 037C 锁存，ELSE 兜底归并 037C（码表声明）；
                  ② 区索引域 0..3 由常量数组界结构性限定，无越界路径（头注释自证）；
                  ③ 故障相挡板输出全保持抬起（安全侧：不拦料）；
                  ④ 无 GVL 依赖：纯引脚输入输出，无外部变量引用，无物理 IO 地址。
  依赖 Depends  : Standard.library（TON / R_TRIG）
  码表 Error codes（Process 段 0005，窗口 037C~037E / 04A4~04A6）:
    16#0005_037C 故障级：组态非法（任一时间域非法）或相位落 ELSE 兜底（归并声明），锁存至 bReset
    16#0005_037D 故障级：释放相单区放行超时（tZoneTo），锁存至 bReset
    16#0005_037E 故障级：积放相满载滞留超时（tAccumTo），锁存至 bReset
    16#0005_04A4 信息级：放行序列启动沿（进 eRel）
    16#0005_04A5 信息级：单区放行完成沿（区光电放空拍）
    16#0005_04A6 信息级：全区放行完成沿（回 eIdle）
  修订历史 Revision :
    2026-11-19  v1.0.0  R42 首版（批次 1 · 序号 5）
*)

TYPE E_DL_GfaState :
(
    eIdle   := 0,    // 积放保持：挡板抬起拦料 / Accum hold, stoppers up
    eRel    := 10,   // 放行：逐区落板放空 / Release, zone-by-zone pass
    eFault  := 90    // 故障：超时锁定 / Fault, latched
);
END_TYPE

FUNCTION_BLOCK FB_DL_GlassFeederAccum
VAR_INPUT
    a_bZonePE    : ARRAY[0..3] OF BOOL;  // 4 区光电，TRUE = 区内有料 [-] / Zone photoeyes, TRUE = occupied
    bConvRun     : BOOL := FALSE;        // 输送运行反馈（当拍量）[-] / Conveyor running feedback
    bRelCmd      : BOOL := FALSE;        // 放行指令，上升沿启动释放序列 [-] / Release command edge
    tZoneTo      : TIME := T#8S;         // 单区放行超时 [ms]，域 > 0 / Per-zone release timeout
    tAccumTo     : TIME := T#60S;        // 满载滞留超时 [ms]，域 > 0 / Full-load dwell timeout
    bReset       : BOOL := FALSE;        // 复位，上升沿清故障锁存 / Reset edge clears fault latch
END_VAR
VAR_OUTPUT
    eState       : E_DL_GfaState;     // 状态出口，段尾单点映射 / State outlet
    a_bStopperUp : ARRAY[0..3] OF BOOL;   // 4 区挡板抬起指令，TRUE = 拦料 [-] / Stopper-up commands
    nRelZone     : DINT;              // 当前放行区号 [0..3]，-1 = 非放行相 / Current releasing zone
    bError       : BOOL;              // 故障锁存标志 / Fault latch flag
    nErrId       : UDINT;             // 事件码，0 = 无事件 / Event code
END_VAR
VAR
    tonZoneTo    : TON;               // 单区放行超时（单相独占），无条件刷新 / Zone release timeout
    tonAccumTo   : TON;               // 满载滞留超时（电平式），无条件刷新 / Full-load dwell timeout
    rtRelCmd     : R_TRIG;            // 放行指令沿实例，无条件刷新 / Release edge instance
    rtReset      : R_TRIG;            // 复位沿实例，无条件刷新 / Reset edge instance
    _eState      : E_DL_GfaState := E_DL_GfaState.eIdle;  // 内部相位（CASE 唯一写入目标）/ Internal phase
    _nRelZoneIdx : DINT := 0;         // 放行序列区号游标 [0..3] / Release sequence zone cursor
    _nIdx        : DINT;              // 阵列循环索引 [-] / Array loop index
    _bAllFull    : BOOL;              // 全区占满当拍量 [-] / All-zones-full current-scan flag
    _bFault      : BOOL;              // 故障锁存位（锁存量）/ Latched fault bit
    _uFault      : UDINT;             // 故障码锁存（锁存量）/ Latched fault code
    _uInfo       : UDINT;             // 信息码，每拍重算 / Transient info code
END_VAR

(* —— 段 0：定时器与沿实例无条件周期刷新（禁置于 IF/CASE 内） —— *)
_bAllFull := a_bZonePE[0] AND a_bZonePE[1] AND a_bZonePE[2] AND a_bZonePE[3];
                                        // 全区占满（当拍量，展开式判据）
rtRelCmd(CLK := bRelCmd);               // 放行沿（每拍必调）
rtReset(CLK := bReset);                 // 复位沿（每拍必调）
tonZoneTo(IN := (_eState = E_DL_GfaState.eRel), PT := tZoneTo);
                                        // 单区放行超时（释放相独占，跨相 IN 必断）
tonAccumTo(IN := (_eState = E_DL_GfaState.eIdle) AND bConvRun AND _bAllFull, PT := tAccumTo);
                                        // 满载滞留超时（电平式，任一条件消失自动断 IN）

(* —— 段 1：单拍量预清零（锁存量 _bFault/_uFault 不入清单，禁同拍抹除） —— *)
_uInfo := 16#0000_0000;             // 信息码每拍重算
nRelZone := -1;                     // 放行区号缺省 -1 = 非放行相
nErrId := 16#0000_0000;             // 事件码缺省无事件

(* —— 段 2：复位沿 + 组态域闸（当拍量判据） —— *)
IF rtReset.Q THEN                   // rtReset.Q = 当拍量
    _bFault := FALSE;               // 清故障锁存位
    _uFault := 16#0000_0000;        // 清故障锁存码
END_IF
IF (TIME_TO_DINT(tZoneTo) <= 0) OR (TIME_TO_DINT(tAccumTo) <= 0) THEN
    _uFault := 16#0005_037C;        // 故障级：组态非法
    _bFault := TRUE;                // 故障标志与码位配对（R45）
END_IF

(* —— 段 3：释放相超时与满载滞留锁存（判据当拍量/单相独占 TON） —— *)
IF (NOT _bFault) AND tonZoneTo.Q THEN
    _uFault := 16#0005_037D;        // 故障级：单区放行超时
    _bFault := TRUE;
END_IF
IF (NOT _bFault) AND tonAccumTo.Q THEN
    _uFault := 16#0005_037E;        // 故障级：满载滞留超时
    _bFault := TRUE;
END_IF

(* —— 段 4：故障解除式（R240 落地，逐 BOOL 标注）：
     rtReset.Q = 当拍量；NOT bRelCmd = 当拍量；a_bZonePE 各元素 = 当拍量。
     均不含锁存量（_bFault/_uFault），解除边真实可达（料清空 + 指令撤销 + 复位沿）。 —— *)
IF rtReset.Q AND (NOT bRelCmd)
   AND (NOT a_bZonePE[0]) AND (NOT a_bZonePE[1])
   AND (NOT a_bZonePE[2]) AND (NOT a_bZonePE[3]) THEN
    _bFault := FALSE;               // 清故障锁存位（锁存量，仅此当拍量解除沿可清）
    _uFault := 16#0000_0000;        // 清故障锁存码（锁存量，仅本当拍量解除沿可清）
    IF _eState = E_DL_GfaState.eFault THEN
        _eState := E_DL_GfaState.eIdle;     // 故障相迁出：回积放保持
    END_IF
END_IF

(* —— 段 5：相位机（CASE 全覆盖 + ELSE 兜底） —— *)
CASE _eState OF

E_DL_GfaState.eIdle:
    FOR _nIdx := 0 TO 3 DO              // 挡板全抬起（拦料保持）
        a_bStopperUp[_nIdx] := TRUE;    // 抬板指令
    END_FOR
    IF rtRelCmd.Q AND (NOT _bFault) THEN
        _nRelZoneIdx := 0;              // 放行游标自下游区 0 起
        _uInfo := 16#0005_04A4;         // 信息级：放行序列启动沿
        _eState := E_DL_GfaState.eRel;  // 进放行相（自区 0 起）
    END_IF

E_DL_GfaState.eRel:
    nRelZone := _nRelZoneIdx;           // 当前放行区号镜像
    a_bStopperUp[_nRelZoneIdx] := FALSE;    // 落板放行当前区
    IF NOT a_bZonePE[_nRelZoneIdx] THEN // 当前区光电放空（当拍量）
        a_bStopperUp[_nRelZoneIdx] := TRUE;     // 抬板恢复拦截
        _uInfo := 16#0005_04A5;         // 信息级：单区放行完成沿
        _nRelZoneIdx := _nRelZoneIdx + 1;       // 进下一区
        IF _nRelZoneIdx > 3 THEN        // 全区放空（索引域 0..3 上界结构性安全）
            _uInfo := 16#0005_04A6;     // 信息级：全区放行完成沿
            _eState := E_DL_GfaState.eIdle;     // 回积放保持相
        END_IF
    END_IF
    (* 超时迁出在段 3 承载 *)

E_DL_GfaState.eFault:
    FOR _nIdx := 0 TO 3 DO              // 故障相挡板全抬起（安全侧：不拦料）
        a_bStopperUp[_nIdx] := TRUE;    // 抬板指令
    END_FOR

ELSE
    _uFault := 16#0005_037C;            // 故障级：非法相位兜底（归并组态码，码表声明）
    _bFault := TRUE;
    _eState := E_DL_GfaState.eFault;    // 强制回故障相

END_CASE

(* —— 段 6：出口单点映射（名实同源；锁存码回放，禁同拍抹除） —— *)
IF _bFault THEN
    nErrId := _uFault;              // 故障锁存码回放
    nRelZone := -1;                 // 故障相放行区号恢复非放行哨兵
ELSE
    nErrId := _uInfo;               // 信息码
END_IF
bError := _bFault;                  // 故障标志与锁存位同源
eState := _eState;                  // 状态出口单点映射

END_FUNCTION_BLOCK

(* ---- FB_DL_GowningRoomSeq.st ---- *)
(*
  ==================================================================
  组件名 Component  : FB_DL_GowningRoomSeq
  分类   Category   : DL_Process
  复杂度 Complexity  : cx5
  版本   Version    : 1.0.0
  功能   Purpose    : 洁净室更衣室顺控。进入请求 → 开入侧门（人进 + 门关反
                      馈）→ 更衣中（完成信号或时限）→ 开出侧门（人出 + 门
                      关反馈）→ 回空闲。双门互锁绝不同开（双命令硬互锁）；
                      更衣时限超时判故障；与 AirShowerInterlockSeq /
                      PassboxInterlockSeq 构成人流三件（ROADMAP 1087 行）。
  来源   Source     : roadmap-p2（R56 评估项落地）
  溯源   Origin     : IEC 61131-3 标准语义的道莅防御性实现；更衣室双门互锁
                      为公开洁净室工艺语义，clean-room 自研实现，未复制任何
                      厂商私有库源码。
  平台   Platform   : 纯 IEC 61131-3（Standard.library: TON / R_TRIG，无私有库）
  分工声明 Split     : 与 FB_DL_AirShowerInterlockSeq 分工——风淋件做吹扫除
                      尘互锁，本件只做更衣流程双门顺控；与
                      FB_DL_PassboxInterlockSeq 分工——传递窗做物件传递，
                      本件做人员进出，两者门数与传感语义不同。
  作者   Author     : 道莅代码库 · PLC 编程专家（R58）
  ------------------------------------------------------------------
  边界 Boundary     :
                      一 双门硬互锁：bDoorInCmd 与 bDoorOutCmd 互为反闸（统
                         一出口单点映射保证绝不同时为真，命令级互锁）；
                      二 更衣时限 tGownMax（执行相看门狗，使能只用相驻留
                         R145）；超时判故障级锁存，双门命令安全侧全断；
                      三 等待类相退出条件 ≥2（R98）：eEnterExit 相 = 人出
                         检测沿或门关反馈（事件）+ 门关前置消失；eChanging
                         相 = 更衣完成信号（事件）+ 时限超时（前置消失）；
                      四 门确认窗配比约束（R100）：tDoorConfirm < tGownMax；
                         越域判故障级；
                      五 故障锁存解除路径 = bReset 上升沿（唯一路径，R188）；
                      六 无全局变量、无外部变量声明、无物理地址寻址。
  修订记录 Revision  :
    2026-11-21  v1.0.0  R58 首版（批 4 · 序号 14）
  ==================================================================
*)

TYPE E_DL_GrpPhase :
(
    eGrpIdle    := 0,  // 空闲：双门关闭等请求 / idle, both doors closed
    eGrpEnter   := 10, // 进入：入侧门开，等人进且门关 / entering, the inner door open
    eGrpChanging:= 20, // 更衣中：双门全闭，等完成信号或时限 / changing, both doors closed
    eGrpExit    := 30, // 离开：出侧门开，等人出且门关 / exiting, the outer door open
    eGrpFault   := 90  // 故障锁存 / the latched fault
);
END_TYPE

TYPE E_DL_GrpFault :
(
    eNone         := 0, // 无成因 / no cause
    eCfgBad       := 1, // 组态非法：门确认窗与更衣时限配比越域（故障级，与 bError 配对）/ an illegal config
    eDoorInTo     := 2, // 入侧门确认超时（故障级，与 bError 配对）/ an inner door confirm timeout
    eGownTimeout  := 3, // 更衣时限超时（故障级，与 bError 配对）/ a gowning timeout
    eDoorOutTo    := 4, // 出侧门确认超时（故障级，与 bError 配对）/ an outer door confirm timeout
    ePhaseBad     := 5  // 非法相位兜底（故障级，与 bError 配对）/ an illegal phase fallback
);
END_TYPE

FUNCTION_BLOCK FB_DL_GowningRoomSeq
VAR_INPUT
    bEnable      : BOOL := TRUE;   // 使能，失能回空闲双门关 [-] / enable, disabling returns idle with both doors closed
    bReset       : BOOL := FALSE;  // 复位上升沿清故障锁存 [-] / reset rising edge clears the latch
    bReqEnter    : BOOL := FALSE;  // 进入请求电平 [-] / the enter request level
    bDoorInClosed: BOOL := TRUE;   // 入侧门关到位反馈 [-] / the inner door closed feedback
    bDoorOutClosed: BOOL := TRUE;  // 出侧门关到位反馈 [-] / the outer door closed feedback
    bPersonIn    : BOOL := FALSE;  // 室内有人检测（更衣室内）[-] / the person inside detection
    bGownDone    : BOOL := FALSE;  // 更衣完成信号（更衣室按钮或工装传感）[-] / the gowning done signal
    tDoorConfirm : TIME := T#10S;  // 门开确认窗 [毫秒] / the door confirm window [millisecond]
    tGownMax     : TIME := T#300S; // 更衣时限 [毫秒] / the gowning max duration [millisecond]
END_VAR
VAR_OUTPUT
    bDoorInCmd : BOOL := FALSE; // 入侧门开门命令输出 [-] / the inner door open command outlet
    bDoorOutCmd: BOOL := FALSE; // 出侧门开门命令输出 [-] / the outer door open command outlet
    bChanging  : BOOL := FALSE; // 更衣进行指示 [-] / the changing indicator
    ePhase     : E_DL_GrpPhase := E_DL_GrpPhase.eGrpIdle; // 相位出口 [枚举] / the phase outlet
    eFault     : E_DL_GrpFault := E_DL_GrpFault.eNone; // 成因出口，锁存回放 [枚举] / the cause outlet replayed
    bError     : BOOL := FALSE; // 故障锁存标志 [-] / the fault latch flag
END_VAR
VAR
    rtReset : R_TRIG; // 复位沿检测，段 0 无条件刷新 / the reset edge
    tonDoor : TON;    // 门开确认窗，段 0 无条件刷新（入 / 出两相共用，相闸区分）/ the door confirm window shared by both door phases
    tonGown : TON;    // 更衣时限窗，段 0 无条件刷新 / the gowning max window
    _ePhase : E_DL_GrpPhase := E_DL_GrpPhase.eGrpIdle; // 内部相位，CASE 唯一写入目标 / the internal phase
    _eFaulC : E_DL_GrpFault := E_DL_GrpFault.eNone; // 故障级成因，锁存至复位沿 / the fault cause latched
    _bFault : BOOL := FALSE; // 故障锁存位 [-] / the fault latch bit
    _bCfgOk : BOOL := FALSE; // 组态域内 [-] / the config inside the domain
    _bInit  : BOOL := FALSE; // 首扫初始化完成标志（R310）/ the first scan flag
END_VAR

// 段 0｜定时器与沿检测无条件周期刷新（禁入分支，FB50-1）/ segment 0, the unconditional refresh
rtReset(CLK := bReset); // 复位沿 / the reset edge
tonDoor(IN := ((_ePhase = E_DL_GrpPhase.eGrpEnter) OR (_ePhase = E_DL_GrpPhase.eGrpExit)) AND (NOT _bFault) AND bEnable, PT := tDoorConfirm); // 门确认窗，IN 串两个开门相闸 / the door window gated by the two open phases
tonGown(IN := (_ePhase = E_DL_GrpPhase.eGrpChanging) AND (NOT _bFault) AND bEnable, PT := tGownMax); // 更衣时限窗，IN 串更衣相闸（纯相驻留，R145）/ the gown window gated by the changing phase

// 段 1｜首扫初始化（R310）/ segment 1, the first scan
IF NOT _bInit THEN // 首扫一拍 / the first scan
    _bInit := TRUE; // 置首扫标志 / raise the flag
END_IF

// 段 2｜复位沿作用域：清故障锁存 / 迁空闲（两项逐项声明，边界五）/ segment 2, the reset edge scope
IF rtReset.Q THEN // 复位沿 / the reset edge
    _bFault := FALSE; // 作用域一：清故障锁存 / scope one, clear the fault latch
    _eFaulC := E_DL_GrpFault.eNone; // 作用域一：清成因 / scope one, clear the cause
    _ePhase := E_DL_GrpPhase.eGrpIdle; // 作用域二：迁空闲相 / scope two, back to idle
END_IF

// 段 3｜组态域闸（边界四，R100 配比：门确认窗 < 更衣时限）/ segment 3, the config gate
_bCfgOk := (tDoorConfirm > T#0S) AND (tGownMax > tDoorConfirm); // 确认窗域与配比判定 / the window domain and the pairing verdict
IF NOT _bCfgOk THEN // 配比越域 / a pairing violation
    IF NOT _bFault THEN // 未锁存才迁移 / migrate only while unlatched
        _bFault := TRUE; // 置故障锁存 / raise the fault latch
        _eFaulC := E_DL_GrpFault.eCfgBad; // 故障级成因（R45 配对）/ the fault cause
        _ePhase := E_DL_GrpPhase.eGrpFault; // 迁故障相（锁存与迁相同分支，FB50-1）/ migrate to the fault phase
    END_IF
END_IF

// 段 4｜相位机：ENUM + CASE，含 ELSE 非法相位兜底（R128）/ segment 4, the phase machine
CASE _ePhase OF

E_DL_GrpPhase.eGrpIdle: // 空闲相：等进入请求（双门关反馈一致性预检）/ the idle phase, awaiting the enter request
    IF NOT bEnable THEN // 失能驻留 / dwell while disabled
        _ePhase := E_DL_GrpPhase.eGrpIdle; // 停摆驻留 / dwell
    ELSIF bReqEnter AND bDoorInClosed AND bDoorOutClosed AND (NOT _bFault) THEN // 请求且双门关确认 / a request with both doors confirmed closed
        _ePhase := E_DL_GrpPhase.eGrpEnter; // 迁进入相 / migrate to the enter phase
    END_IF

E_DL_GrpPhase.eGrpEnter: // 进入相：入侧门开，等人进且门关（R98 事件 + 前置消失）/ the enter phase
    IF NOT bEnable THEN // 失能回空闲 / a disable returns idle
        _ePhase := E_DL_GrpPhase.eGrpIdle; // 回空闲相 / back to idle
    ELSIF bPersonIn AND bDoorInClosed THEN // 人进且入侧门关（事件与前置消失双条件）/ the person in with the door closed
        _ePhase := E_DL_GrpPhase.eGrpChanging; // 迁更衣相 / migrate to the changing phase
    ELSIF tonDoor.Q THEN // 门确认窗超时（R190 独立成因）/ the door confirm timeout, an independent cause
        _bFault := TRUE; // 置故障锁存 / raise the fault latch
        _eFaulC := E_DL_GrpFault.eDoorInTo; // 故障级成因（R45 配对）/ the fault cause
        _ePhase := E_DL_GrpPhase.eGrpFault; // 迁故障相 / migrate to the fault phase
    END_IF

E_DL_GrpPhase.eGrpChanging: // 更衣相：双门全闭，等完成信号或时限（边界三双出口）/ the changing phase, the dual exit
    IF NOT bEnable THEN // 失能回空闲（R191 显式：门命令安全侧全断）/ a disable returns idle
        _ePhase := E_DL_GrpPhase.eGrpIdle; // 回空闲相 / back to idle
    ELSIF bGownDone THEN // 更衣完成信号（事件）/ the gowning done event
        _ePhase := E_DL_GrpPhase.eGrpExit; // 迁离开相 / migrate to the exit phase
    ELSIF tonGown.Q THEN // 更衣时限超时（前置消失路径，R190 独立成因）/ the gown timeout, the precondition lost path
        _bFault := TRUE; // 置故障锁存 / raise the fault latch
        _eFaulC := E_DL_GrpFault.eGownTimeout; // 故障级成因（R45 配对）/ the fault cause
        _ePhase := E_DL_GrpPhase.eGrpFault; // 迁故障相 / migrate to the fault phase
    END_IF

E_DL_GrpPhase.eGrpExit: // 离开相：出侧门开，等人出且门关 / the exit phase
    IF NOT bEnable THEN // 失能回空闲 / a disable returns idle
        _ePhase := E_DL_GrpPhase.eGrpIdle; // 回空闲相 / back to idle
    ELSIF (NOT bPersonIn) AND bDoorOutClosed THEN // 人出且出侧门关 / the person out with the door closed
        _ePhase := E_DL_GrpPhase.eGrpIdle; // 回空闲相 / back to idle
    ELSIF tonDoor.Q THEN // 门确认窗超时（R190 独立成因）/ the door confirm timeout
        _bFault := TRUE; // 置故障锁存 / raise the fault latch
        _eFaulC := E_DL_GrpFault.eDoorOutTo; // 故障级成因（R45 配对）/ the fault cause
        _ePhase := E_DL_GrpPhase.eGrpFault; // 迁故障相 / migrate to the fault phase
    END_IF

E_DL_GrpPhase.eGrpFault: // 故障相：成因锁存等复位沿；双门命令安全侧全断 / the fault phase
ELSE // 非法相位兜底（R128）/ the illegal phase fallback
    _bFault := TRUE; // 置故障锁存 / raise the fault latch
    _eFaulC := E_DL_GrpFault.ePhaseBad; // 故障级成因（R45 配对）/ the fault cause
    _ePhase := E_DL_GrpPhase.eGrpFault; // 迁故障相 / migrate to the fault phase
END_CASE

// 段 5｜统一出口：双门互锁单点映射（边界一）/ segment 5, the unified outlet with the interlock
bDoorInCmd := (_ePhase = E_DL_GrpPhase.eGrpEnter) AND bEnable AND (NOT _bFault); // 入侧命令仅进入相（互锁）/ the inner command in the enter phase only
bDoorOutCmd := (_ePhase = E_DL_GrpPhase.eGrpExit) AND bEnable AND (NOT _bFault); // 出侧命令仅离开相（互锁）/ the outer command in the exit phase only
bChanging := _ePhase = E_DL_GrpPhase.eGrpChanging; // 更衣指示 / the changing indicator
ePhase := _ePhase; // 相位出口单点映射 / the phase outlet
IF _bFault THEN // 故障锁存优先 / the fault latch first
    eFault := _eFaulC; // 成因锁存回放（R152）/ the cause replayed
ELSE // 无锁存 / no latch
    eFault := E_DL_GrpFault.eNone; // 无成因 / no cause
END_IF
bError := _bFault; // 故障标志与锁存位同源 / the flag shares the latch
END_FUNCTION_BLOCK
